(* IEC 61131-3 sources: daoli-st-library/DL_Process (part 42) *)

(* ---- FB_DL_MoldingLineSandSeq.st ---- *)
(*
 * FB_DL_MoldingLineSandSeq | C4 | DL_Process
 * 功能：造型线「回砂→磁选→冷却→混砂→松砂→造型→浇注」序列控制；每相独立使能出口 + 独立 TON 超时，冷却相按砂温判据转出、浇注相按许可驻留       单位：温度 [℃]、rTimeoutS [s]、码位 [INT]
 * 工况边界：COOLING 只在 rSandTempC ≤ rSandTempMaxC 时转 MULLING，超时判 9701；POURING 无 xPourPermit 时驻留并只发告警 9702（告警级，不置 xFault），浇注相超时判 9709；砂温 NaN/±Inf 或越量程（-20~200 ℃）判 9708；rTimeoutS 须 >0；xStart 只用上升沿启动，xStop 按逆序（浇注→造型→松砂→混砂→冷却→磁选→回砂）撤令
 * 代数值回代：rSandTempC=42.0 ≤ rSandTempMaxC=45 → 冷却完成转混砂；rSandTempC=52.0 >45 → 驻留冷却直至 9701（与 spec 判据一致）
 * 开源溯源：clean-room 自研，未复制任何第三方代码（无外部来源）
 *)
(*
 * 码位总账（本件故障码全清单，逐条在实现分支中可到达；故障级锁存回放）：
 * 9701 冷却温度超时 / 9702 浇注许可缺失（告警级，不置 xFault）/ 9703 回砂相就绪丢失 / 9704 磁选相回砂就绪丢失 / 9705 混砂相供砂就绪丢失 / 9706 松砂相造型机未就绪 / 9707 造型相就绪未建立 / 9708 砂温或参数非法 / 9709 浇注超时（故障锁存，清除沿 = xStart 下降沿）；MAGNET/MULLING/AERATING 正常以驻留定时转出，其码位仅在就绪丢失时置位
 *)

TYPE E_DL_SandLinePhase :
(
    IDLE        := 0,    // 待机，全部命令撤销 | idle, every command withdrawn
    RETURN_SAND := 10,   // 回砂相，旧砂输送 | return sand conveying
    MAGNET      := 20,   // 磁选相，除铁器投入 | magnetic separation
    COOLING     := 30,   // 冷却相，沸腾冷却床 | cooling bed
    MULLING     := 40,   // 混砂相，混砂机加水加膨润土 | mulling
    AERATING    := 50,   // 松砂相，松砂机打散 | aerating
    MOLDING     := 60,   // 造型相，造型机射砂压实 | molding
    POURING     := 70,   // 浇注相，等待浇注许可 | pouring, waiting for the permit
    FAULT       := 90    // 故障相，全部命令强制 FALSE，码位锁存 | fault phase, all commands forced FALSE, the code is latched
);
END_TYPE

FUNCTION_BLOCK FB_DL_MoldingLineSandSeq
VAR_INPUT
    xStart        : BOOL;            // 启动（下降沿兼作故障复位沿）| start, its falling edge also resets a latched fault
    xStop         : BOOL;            // 停止（任意相生效，逆序停车）| stop, effective in any phase and stopping in reverse order
    xSandReady    : BOOL;            // 回砂段就绪 | return sand section ready
    xMoldReady    : BOOL;            // 造型机就绪 | molding machine ready
    xPourPermit   : BOOL;            // 浇注许可（来自浇注机/行车）| pouring permit from the pouring device
    rSandTempC    : REAL;            // 型砂温度 | molding sand temperature [℃]
    rSandTempMaxC : REAL := 45.0;    // 允许混砂的最高砂温 | maximum sand temperature for mulling [℃]
    rTimeoutS     : REAL := 90.0;    // 每相超时设定 | per-phase timeout setting [s]
END_VAR
VAR_OUTPUT
    xReturnCmd : BOOL;               // 回砂命令（RETURN_SAND 相独立使能）| return sand command, independent enable
    xMagnetCmd : BOOL;               // 磁选命令（MAGNET 相独立使能）| magnet command, independent enable
    xCoolCmd   : BOOL;               // 冷却命令（COOLING 相独立使能）| cooling command, independent enable
    xMullerCmd : BOOL;               // 混砂命令（MULLING 相独立使能）| mulling command, independent enable
    xAerateCmd : BOOL;               // 松砂命令（AERATING 相独立使能）| aerating command, independent enable
    xMoldCmd   : BOOL;               // 造型命令（MOLDING 相独立使能）| molding command, independent enable
    xPourCmd   : BOOL;               // 浇注命令（POURING 相且许可到位独立使能）| pouring command, independent enable when permitted
    ePhase     : E_DL_SandLinePhase; // 当前相 | current phase
    xFault     : BOOL;               // 故障标志（仅故障级码置位）| fault flag, fault-class codes only
    nFaultCode : INT;                // 故障码，锁存至复位沿 | fault code latched until the reset edge
    nWarnCode  : INT;                // 告警码（9702 浇注许可缺失，信息级不置 xFault）| warning code for the missing pouring permit
END_VAR
VAR
    tonReturn : TON;                 // RETURN_SAND 相超时定时器 | timeout of RETURN_SAND
    tonMagnet : TON;                 // MAGNET 相超时定时器 | timeout of MAGNET
    tonCool   : TON;                 // COOLING 相超时定时器 | timeout of COOLING
    tonMull   : TON;                 // MULLING 相超时定时器 | timeout of MULLING
    tonAerate : TON;                 // AERATING 相超时定时器 | timeout of AERATING
    tonMold   : TON;                 // MOLDING 相超时定时器 | timeout of MOLDING
    tonPour   : TON;                 // POURING 相超时定时器 | timeout of POURING
    fbStartRise : R_TRIG;            // xStart 上升沿（唯一启动沿）| rising edge of xStart, the single start edge
    fbStartFall : F_TRIG;            // xStart 下降沿（故障复位沿）| falling edge of xStart, the fault reset edge
    xParamOk  : BOOL;                // 超时与砂温上限参数合法 | timeout and sand temperature limit are legal
    xFinTemp  : BOOL;                // 砂温有限性 | sand temperature is finite
    xTempBad  : BOOL;                // 砂温非有限或越量程 | sand temperature non-finite or out of range
    xCoolDone : BOOL;                // 冷却到位（砂温 ≤ 上限）| cooling done, temperature within the limit
    nTmoMs    : UDINT := 90000;      // 超时毫秒数（缺省值防首拍 PT=0 假超时）| timeout in milliseconds, default prevents a zero PT
    nCodeLatch: INT;                 // 故障码锁存副本 | latched copy of the fault code
END_VAR
VAR CONSTANT
    DL_SLS_TEMP_MAX : REAL := 200.0; // 砂温量程上限 | upper sand temperature limit [℃]
    DL_SLS_TEMP_MIN : REAL := -20.0; // 砂温量程下限 | lower sand temperature limit [℃]
    DL_SLS_C_COOL   : INT := 9701;   // 冷却温度超时 | cooling temperature timeout
    DL_SLS_C_PERMIT : INT := 9702;   // 浇注许可缺失（告警级）| missing pouring permit, warning class
    DL_SLS_C_RETURN : INT := 9703;   // 回砂超时 | return sand timeout
    DL_SLS_C_MAGNET : INT := 9704;   // 磁选超时 | magnet timeout
    DL_SLS_C_MULL   : INT := 9705;   // 混砂超时 | mulling timeout
    DL_SLS_C_AERATE : INT := 9706;   // 松砂超时 | aerating timeout
    DL_SLS_C_MOLD   : INT := 9707;   // 造型超时 | molding timeout
    DL_SLS_C_BAD    : INT := 9708;   // 砂温或参数非法 | sand temperature or parameter illegal
    DL_SLS_C_POUR   : INT := 9709;   // 浇注超时 | pouring timeout
END_VAR

// 段1｜参数与采样门禁（先判后用：REAL→UDINT 换算在闸后进行，结果供段2 定时器使用）
xParamOk := (rTimeoutS = rTimeoutS) AND ((rTimeoutS - rTimeoutS) = 0.0) AND (rTimeoutS > 0.0)
            AND (rSandTempMaxC = rSandTempMaxC) AND ((rSandTempMaxC - rSandTempMaxC) = 0.0);
IF xParamOk THEN
    nTmoMs := REAL_TO_UDINT(rTimeoutS * 1000.0);
ELSE
    nTmoMs := 90000;                 // 参数非法取保守值 | conservative value on an illegal parameter
END_IF
xFinTemp := (rSandTempC = rSandTempC) AND ((rSandTempC - rSandTempC) = 0.0);
xTempBad := (NOT xFinTemp) OR (rSandTempC > DL_SLS_TEMP_MAX) OR (rSandTempC < DL_SLS_TEMP_MIN);
xCoolDone := (NOT xTempBad) AND (rSandTempC <= rSandTempMaxC);

// 段2｜七只定时器 + 两只边沿实例无条件周期刷新（R7，一相一只实例不跨相复用；PT 取自段1 已换算毫秒值）
tonReturn(IN := ePhase = E_DL_SandLinePhase.RETURN_SAND, PT := UDINT_TO_TIME(nTmoMs));
tonMagnet(IN := ePhase = E_DL_SandLinePhase.MAGNET, PT := UDINT_TO_TIME(nTmoMs));
tonCool(IN := ePhase = E_DL_SandLinePhase.COOLING, PT := UDINT_TO_TIME(nTmoMs));
tonMull(IN := ePhase = E_DL_SandLinePhase.MULLING, PT := UDINT_TO_TIME(nTmoMs));
tonAerate(IN := ePhase = E_DL_SandLinePhase.AERATING, PT := UDINT_TO_TIME(nTmoMs));
tonMold(IN := ePhase = E_DL_SandLinePhase.MOLDING, PT := UDINT_TO_TIME(nTmoMs));
tonPour(IN := ePhase = E_DL_SandLinePhase.POURING, PT := UDINT_TO_TIME(nTmoMs));
fbStartRise(CLK := xStart);
fbStartFall(CLK := xStart);

// 段3｜输出预置（唯一预置点，CASE 内只置位）
xReturnCmd := FALSE;
xMagnetCmd := FALSE;
xCoolCmd := FALSE;
xMullerCmd := FALSE;
xAerateCmd := FALSE;
xMoldCmd := FALSE;
xPourCmd := FALSE;
xFault := FALSE;
nFaultCode := 0;
nWarnCode := 0;

// 段4｜全局闸：参数/砂温非法 → 锁故障；xStop → 逆序停车
IF (NOT xParamOk) OR xTempBad THEN
    nCodeLatch := DL_SLS_C_BAD;
    xFault := TRUE;
    nFaultCode := DL_SLS_C_BAD;
    ePhase := E_DL_SandLinePhase.FAULT;
ELSIF xStop AND (ePhase <> E_DL_SandLinePhase.IDLE) THEN
    xPourCmd := FALSE;               // 逆序停车第 1 步：浇注先停 | reverse stop step 1, pouring first
    xMoldCmd := FALSE;               // 逆序停车第 2 步：造型 | step 2, molding
    xAerateCmd := FALSE;             // 逆序停车第 3 步：松砂 | step 3, aerating
    xMullerCmd := FALSE;             // 逆序停车第 4 步：混砂 | step 4, mulling
    xCoolCmd := FALSE;               // 逆序停车第 5 步：冷却 | step 5, cooling
    xMagnetCmd := FALSE;             // 逆序停车第 6 步：磁选 | step 6, magnet
    xReturnCmd := FALSE;             // 逆序停车第 7 步：回砂最后停（下游优先，同拍置假）| step 7, return sand last
    ePhase := E_DL_SandLinePhase.IDLE;
END_IF

// 段5｜主状态机（ENUM + CASE，ELSE 兜底）
IF ePhase <> E_DL_SandLinePhase.FAULT THEN
CASE ePhase OF
E_DL_SandLinePhase.IDLE:
    // 拍 N：待机，仅 xStart 上升沿且回砂就绪时启动（防停车后自恢复）
    IF fbStartRise.Q AND xSandReady AND (NOT xStop) THEN
        ePhase := E_DL_SandLinePhase.RETURN_SAND;     // 本拍行为：进回砂相 | enter return sand
    END_IF

E_DL_SandLinePhase.RETURN_SAND:
    // 拍 N：回砂输送到位由驻留定时判完成；期间回砂就绪丢失即报 9703（启动条件已含 xSandReady，故不以其为转出条件）
    IF NOT xSandReady THEN
        nCodeLatch := DL_SLS_C_RETURN;                // 回砂就绪丢失 | return sand readiness lost
        xFault := TRUE;
        nFaultCode := DL_SLS_C_RETURN;
        ePhase := E_DL_SandLinePhase.FAULT;
    ELSIF tonReturn.Q THEN
        ePhase := E_DL_SandLinePhase.MAGNET;          // 本拍行为：进磁选相 | enter magnet
    END_IF

E_DL_SandLinePhase.MAGNET:
    // 拍 N：磁选除铁，回砂段中断即报 9704；正常由驻留定时转冷却
    IF NOT xSandReady THEN
        nCodeLatch := DL_SLS_C_MAGNET;                // 回砂段中断，磁选无法维持 | return sand interrupted
        xFault := TRUE;
        nFaultCode := DL_SLS_C_MAGNET;
        ePhase := E_DL_SandLinePhase.FAULT;
    ELSIF tonMagnet.Q THEN
        ePhase := E_DL_SandLinePhase.COOLING;         // 本拍行为：进冷却相 | enter cooling
    END_IF

E_DL_SandLinePhase.COOLING:
    // 拍 N：沸腾冷却，砂温降到上限以下才进混砂；超时判 9701
    IF xCoolDone THEN
        ePhase := E_DL_SandLinePhase.MULLING;         // 本拍行为：砂温达标进混砂 | sand cool enough, enter mulling
    ELSIF tonCool.Q THEN
        nCodeLatch := DL_SLS_C_COOL;                  // 冷却温度超时 | cooling temperature timeout
        xFault := TRUE;
        nFaultCode := DL_SLS_C_COOL;
        ePhase := E_DL_SandLinePhase.FAULT;
    END_IF

E_DL_SandLinePhase.MULLING:
    // 拍 N：混砂（加水、加膨润土），供砂中断即报 9705；正常由驻留定时转松砂
    IF NOT xSandReady THEN
        nCodeLatch := DL_SLS_C_MULL;                  // 供砂中断，混砂配比失真 | sand supply interrupted, the batch would be off-ratio
        xFault := TRUE;
        nFaultCode := DL_SLS_C_MULL;
        ePhase := E_DL_SandLinePhase.FAULT;
    ELSIF tonMull.Q THEN
        ePhase := E_DL_SandLinePhase.AERATING;        // 本拍行为：进松砂相 | enter aerating
    END_IF

E_DL_SandLinePhase.AERATING:
    // 拍 N：松砂打散，造型机未就绪即报 9706（砂无去处）；正常由驻留定时转造型
    IF NOT xMoldReady THEN
        nCodeLatch := DL_SLS_C_AERATE;                // 造型机未就绪，松砂后无处送 | molding machine not ready, no destination
        xFault := TRUE;
        nFaultCode := DL_SLS_C_AERATE;
        ePhase := E_DL_SandLinePhase.FAULT;
    ELSIF tonAerate.Q THEN
        ePhase := E_DL_SandLinePhase.MOLDING;         // 本拍行为：进造型相 | enter molding
    END_IF

E_DL_SandLinePhase.MOLDING:
    // 拍 N：造型射砂压实，等造型机就绪确认与时间窗
    IF tonMold.Q AND xMoldReady THEN
        ePhase := E_DL_SandLinePhase.POURING;         // 本拍行为：进浇注相 | enter pouring
    ELSIF tonMold.Q AND (NOT xMoldReady) THEN
        nCodeLatch := DL_SLS_C_MOLD;                  // 造型就绪始终未建立 | molding readiness never established
        xFault := TRUE;
        nFaultCode := DL_SLS_C_MOLD;
        ePhase := E_DL_SandLinePhase.FAULT;
    END_IF

E_DL_SandLinePhase.POURING:
    // 拍 N：等浇注许可；无许可只驻留并告警 9702，不置故障
    IF NOT xPourPermit THEN
        nWarnCode := DL_SLS_C_PERMIT;                 // 告警级：许可缺失（信息级码永不置 bError）| warning class, never raises the fault flag
        IF tonPour.Q THEN
            nCodeLatch := DL_SLS_C_POUR;              // 浇注超时：锁存 9709 | pouring timeout, latch 9709
            xFault := TRUE;
            nFaultCode := DL_SLS_C_POUR;
            ePhase := E_DL_SandLinePhase.FAULT;
        END_IF
    ELSIF tonPour.Q THEN
        ePhase := E_DL_SandLinePhase.IDLE;            // 本拍行为：浇注完成回待机 | pouring done, back to idle
    END_IF

E_DL_SandLinePhase.FAULT:
    // 故障相（本段被外层 IF 排除，保留分支以满足穷举）
    xFault := TRUE;
    nFaultCode := nCodeLatch;

ELSE
    // 非法状态兜底：绝不停在未知相
    nCodeLatch := DL_SLS_C_BAD;
    xFault := TRUE;
    nFaultCode := DL_SLS_C_BAD;
    ePhase := E_DL_SandLinePhase.FAULT;
END_CASE
END_IF

// 段6｜每相独立使能出口（IDLE/FAULT 不置任何命令，天然强制 FALSE）
CASE ePhase OF
E_DL_SandLinePhase.RETURN_SAND:
    xReturnCmd := TRUE;                           // 回砂相独立使能出口 | independent enable of RETURN_SAND
E_DL_SandLinePhase.MAGNET:
    xMagnetCmd := TRUE;                           // 磁选相独立使能出口 | independent enable of MAGNET
E_DL_SandLinePhase.COOLING:
    xCoolCmd := TRUE;                             // 冷却相独立使能出口 | independent enable of COOLING
E_DL_SandLinePhase.MULLING:
    xMullerCmd := TRUE;                           // 混砂相独立使能出口 | independent enable of MULLING
E_DL_SandLinePhase.AERATING:
    xAerateCmd := TRUE;                           // 松砂相独立使能出口 | independent enable of AERATING
E_DL_SandLinePhase.MOLDING:
    xMoldCmd := TRUE;                             // 造型相独立使能出口 | independent enable of MOLDING
E_DL_SandLinePhase.POURING:
    xPourCmd := xPourPermit;                      // 浇注相独立使能出口（无许可不浇注）| independent enable of POURING, gated by the permit
ELSE
    xReturnCmd := FALSE;                          // 其余相（含 FAULT）：命令强制 FALSE | all other phases force FALSE
    xMagnetCmd := FALSE;
    xCoolCmd := FALSE;
    xMullerCmd := FALSE;
    xAerateCmd := FALSE;
    xMoldCmd := FALSE;
    xPourCmd := FALSE;
END_CASE

// 段7｜故障相锁存回放 + 复位沿（xStart 下降沿清除）
IF ePhase = E_DL_SandLinePhase.FAULT THEN
    xFault := TRUE;
    nFaultCode := nCodeLatch;                     // 锁存回放，不按当下输入重推断 | republish the latch
    xReturnCmd := FALSE;
    xMagnetCmd := FALSE;
    xCoolCmd := FALSE;
    xMullerCmd := FALSE;
    xAerateCmd := FALSE;
    xMoldCmd := FALSE;
    xPourCmd := FALSE;
    nWarnCode := 0;
    IF fbStartFall.Q THEN
        nCodeLatch := 0;                          // 清除边：xStart 下降沿（头注释已声明）| clear edge declared in the header
        ePhase := E_DL_SandLinePhase.IDLE;
    END_IF
END_IF
END_FUNCTION_BLOCK

(* ---- FB_DL_NailMachineSeq.st ---- *)
//==============================================================================
// 功能块：FB_DL_NailMachineSeq ｜ 中文名称：极耳裁切/模切机顺控
// 所属子库：DL_Process ｜ 版本：v1.0.0 ｜ 兼容：CODESYS V3.5+ / TwinCAT 3 / 汇川 InoProShop
// 功能描述：极耳裁切/模切机节拍链——放卷 → 裁切 → 收料三工位联动：
//           三就绪门控起步、单拍节拍超时保护、批量计数达批自动收批；
//           bStop 立即断裁切输出（模切头行程内停止由驱动层负责，边界声明）。
// 开源溯源 (Origin)：道莅原创实现（参考锂电极耳模切机工程惯例 分类与参数域）
// 单位表：计数[片] / 节拍[ms] / 诊断掩码[位]
// 错误码表：16#0005_01E4 信息级（三就绪缺一，诊断掩码输出，不置 bError）/
//           16#0005_01E5 信息级（批量计数达批，正常收批结论，不置 bError）/
//           16#0005_031B 故障级（单拍节拍超时，全停，置 bError）/
//           16#0005_031C 预留禁用（不得挪用）/ 16#0005_031D 故障级兜底
//           （状态机落 ELSE，置 bError 并全停）
// 状态机：E_DL_NailSeqState（七态：eIdle=0 / eWaitReady=10 / eRun=20 /
//           eCutting=30 / eCollecting=40 / eBatchDone=50 / eFault=99），
//           CASE 含 ELSE 兜底，ELSE 置 031D 并全停
// 边界行为：① 三就绪缺一 → 停在 eWaitReady 并输出诊断掩码 uNotReadyMask
//           （位 0 = 放卷缺、位 1 = 裁切原点缺、位 2 = 收料缺）+ 信息 01E4；
//           ② 单拍节拍超时（tCutCycleMax 内未回到原点/收到切完反馈）→
//           故障 031B + 全停；③ 计数达批 → 回 eIdle + 信息 01E5；④ bStop
//           立即断裁切输出（安全侧不停机次序假设：模切头行程内停止由
//           驱动层负责，本件只断输出指令，头注释边界声明）；⑤ 计数饱和
//           4294967295 不回绕；⑥ 非有限/非法防御：批量目标为 0 不判故障
//           （0 = 连续模式），节拍上限 <= 0 判组态非法 031B 复用（R90）。
// 依赖纪律：仅 Standard.library；零跨层调用（三工位节拍编排为自研顺控，
//           不复用 StepSequencer——工位间为并行联动非串行步，复用会扭曲
//           语义，头注释声明此设计取舍）。
// 修订历史：v1.0.0 2026-11-17 首版（R23 派单 · ROADMAP 锂电 P1 §351）
//==============================================================================

(*------------------------------------------------------------------------------
 * 枚举: E_DL_NailSeqState（归属本功能块，同文件发布，全库唯一定义）
 * 含义: 模切机顺控相位，每个成员在 CASE 中有且仅有一个标签。
 *-----------------------------------------------------------------------------*)
TYPE E_DL_NailSeqState :
(
    eIdle       := 0,   // 空闲：等启动 / Idle, awaiting start
    eWaitReady  := 10,  // 等就绪：三工位就绪门控（诊断掩码输出） / Waiting for readiness with a diagnostic mask
    eRun        := 20,  // 运行：放卷 + 收料联动输出 / Running, unwind and collector active
    eCutting    := 30,  // 裁切：切脉冲发出，等切完反馈/回原点 / Cutting, pulse issued, waiting for done or home
    eCollecting := 40,  // 收料：裁切完成转收料拍 / Collecting, the cut done transitions to the collect beat
    eBatchDone  := 50,  // 批完成：达批收批，等启动撤销 / Batch done, awaiting the start drop
    eFault      := 99   // 故障：节拍超时/组态非法/非法状态 / Fault, cycle timeout, illegal config or state
);
END_TYPE

FUNCTION_BLOCK FB_DL_NailMachineSeq
VAR_INPUT
    bStart         : BOOL;                  // 启动请求 [—]，上升沿生效 / Start request, rising edge
    bStop          : BOOL;                  // 停止请求 [—]，电平有效，立即断裁切输出 / Stop request, level active, cut output dropped immediately
    bUnwinderReady : BOOL;                  // 放卷就绪反馈 [—] / Unwinder ready feedback
    bCutterHome    : BOOL;                  // 裁切原点反馈 [—] / Cutter home feedback
    bCollectorReady: BOOL;                  // 收料就绪反馈 [—] / Collector ready feedback
    bCutDone       : BOOL;                  // 切完反馈 [—]，每片一拍 / Cut-done feedback, one scan per piece
    uBatchCount    : UDINT;                 // 批量目标 [片]，0 = 连续模式 / Batch target [pieces], zero = continuous mode
    tCutCycleMax   : TIME := T#3S;          // 单拍节拍上限 [ms]，须 > 0 / Single-cycle ceiling [ms], must be > 0
    bReset         : BOOL;                  // 故障复位 [—]，上升沿退出 eFault / Fault reset, rising edge leaves fault
END_VAR
VAR_OUTPUT
    eSeqState      : E_DL_NailSeqState;     // 顺控相位 [—] / Sequence phase
    uCutDone       : UDINT;                 // 已切计数 [片]，饱和不回绕 / Cut counter [pieces], saturated without wrap
    uNotReadyMask  : UINT;                  // 就绪诊断掩码 [位]，位0放卷/位1原点/位2收料 / Readiness diagnostic mask, bit0 unwind, bit1 home, bit2 collector
    bUnwindRun     : BOOL;                  // 放卷运行输出 [—] / Unwind run output
    bCutTrig       : BOOL;                  // 裁切触发输出 [—] / Cut trigger output
    bCollectRun    : BOOL;                  // 收料运行输出 [—] / Collector run output
    eErr           : UDINT;                 // 错误码，0 = 无错 / Error code, 0 = no error
    bError         : BOOL;                  // 故障级标志，仅故障级错误置位 / Fault-class flag, set only on fault-level codes
    bValid         : BOOL;                  // 输出可用标志 / Outputs usable flag
END_VAR
VAR
    fbCycle        : TON;                   // 单拍节拍计时，段 6 无条件刷新 [ms] / Single-cycle timer
    _eState        : E_DL_NailSeqState := E_DL_NailSeqState.eIdle; // 当前相位 / Current phase
    _bInit         : BOOL := FALSE;         // 首扫标志，初值 FALSE 取非判定 / First-scan flag, tested negated
    _bStartPrev    : BOOL;                  // 启动命令上拍电平快照 / Previous-scan level of the start command
    _bIllegal      : BOOL;                  // 非法状态标志 / Illegal state flag
    _bCfgBad       : BOOL;                  // 组态非法锁存（节拍上限 <= 0） / Illegal configuration latch
    _bNotReady     : BOOL;                  // 三就绪缺一当拍标志 / Readiness-missing flag of this scan
END_VAR
VAR CONSTANT
    DL_NAIL_CNT_MAX : UDINT := 4294967295;  // 计数饱和上限 [片] / Counter saturation ceiling [pieces]
    DL_NAIL_INF     : LREAL := 1.7976931348623157E308; // LREAL 幅值上限（本件无浮点引脚，防御常量备扩展） / LREAL ceiling reserved for extensions
END_VAR

(*------------------------------------------------------------------------------
 * 段 1｜每拍预置：三输出先全断（安全侧），单拍标志预清零
 *      Three outputs cleared first, fail-safe, one-shot flags pre-cleared
 *-----------------------------------------------------------------------------*)
bUnwindRun    := FALSE;                     // 放卷输出先清（安全侧） / Unwind output cleared first
bCutTrig      := FALSE;                     // 裁切输出先清（安全侧） / Cut output cleared first
bCollectRun   := FALSE;                     // 收料输出先清（安全侧） / Collector output cleared first
eErr          := 16#0000_0000;              // 错误码每拍重算 / Error code recomputed
bError        := FALSE;                     // 故障标志每拍重算 / Fault flag recomputed
bValid        := FALSE;                     // 可用标志每拍重算 / Usable flag recomputed
_bIllegal     := FALSE;                     // 非法状态标志预清零 / Illegal flag pre-cleared
_bNotReady    := FALSE;                     // 就绪缺一标志预清零 / Readiness flag pre-cleared
uNotReadyMask := 0;                         // 诊断掩码每拍重算 / Diagnostic mask recomputed

(*------------------------------------------------------------------------------
 * 段 2｜首扫初始化
 *      First-scan initialisation
 *-----------------------------------------------------------------------------*)
IF NOT _bInit THEN
    _eState     := E_DL_NailSeqState.eIdle; // 相位空闲起步 / Phase starts idle
    uCutDone    := 0;                       // 计数清零 / Counter cleared
    _bCfgBad    := FALSE;                   // 组态锁存清零 / Config latch cleared
    _bInit      := TRUE;                    // 首扫只做一次 / The first scan runs once
END_IF

(*------------------------------------------------------------------------------
 * 段 3｜组态闸门：节拍上限 <= 0 → 组态非法（031B 复用，R90）
 *      Configuration gate: non-positive cycle ceiling is illegal
 *-----------------------------------------------------------------------------*)
IF TIME_TO_DINT(tCutCycleMax) <= 0 THEN
    _bCfgBad := TRUE;                       // 组态非法锁存 / Illegal configuration latched
END_IF

(*------------------------------------------------------------------------------
 * 段 4｜就绪门控与诊断掩码装配
 *      Readiness gating and the diagnostic mask assembly
 *-----------------------------------------------------------------------------*)
IF (NOT bUnwinderReady) OR (NOT bCutterHome) OR (NOT bCollectorReady) THEN
    _bNotReady := TRUE;                     // 三就绪缺一 / Readiness missing
    IF NOT bUnwinderReady THEN
        uNotReadyMask := uNotReadyMask OR 1; // 位 0：放卷缺 / Bit 0, unwind missing
    END_IF
    IF NOT bCutterHome THEN
        uNotReadyMask := uNotReadyMask OR 2; // 位 1：裁切原点缺 / Bit 1, home missing
    END_IF
    IF NOT bCollectorReady THEN
        uNotReadyMask := uNotReadyMask OR 4; // 位 2：收料缺 / Bit 2, collector missing
    END_IF
END_IF

(*------------------------------------------------------------------------------
 * 段 5｜单拍节拍计时无条件刷新（R40：CASE 之外每拍必调）
 *      Cycle timer refreshed unconditionally per R40
 *-----------------------------------------------------------------------------*)
fbCycle(IN := (_eState = E_DL_NailSeqState.eCutting), PT := tCutCycleMax); // 单拍节拍计时 / Single-cycle timer

(*------------------------------------------------------------------------------
 * 段 6｜相位机（只做迁移；输出在段 7 按相置位）
 *      Phase machine, transitions only, outputs assigned in segment seven
 *-----------------------------------------------------------------------------*)
CASE _eState OF

    E_DL_NailSeqState.eIdle:               // 空闲：启动沿进等就绪
        IF bStart AND (NOT _bStartPrev) AND (NOT _bCfgBad) THEN
            _eState := E_DL_NailSeqState.eWaitReady; // 进等就绪 / To the wait-ready phase
        END_IF

    E_DL_NailSeqState.eWaitReady:          // 等就绪：三就绪全满进运行
        IF _bNotReady THEN
            _eState := E_DL_NailSeqState.eWaitReady; // 缺一滞留（掩码在段 7 输出） / Held while missing, the mask is output
        ELSE
            _eState := E_DL_NailSeqState.eRun; // 就绪全满，进运行 / All ready, run
        END_IF
        IF bStop THEN
            _eState := E_DL_NailSeqState.eIdle; // 停止请求回空闲 / Stop back to idle
        END_IF

    E_DL_NailSeqState.eRun:                // 运行：放卷 + 收料联动，发裁切触发
        IF bStop OR _bNotReady THEN
            _eState := E_DL_NailSeqState.eIdle; // 停止或缺就绪回空闲 / Stop or missing readiness back to idle
        ELSIF (bCutDone OR NOT bCutterHome) THEN
            _eState := E_DL_NailSeqState.eCutting; // 发切（反馈或离原点即视为切入） / To cutting
        END_IF

    E_DL_NailSeqState.eCutting:            // 裁切：等切完反馈或节拍超时
        IF bStop THEN
            _eState := E_DL_NailSeqState.eIdle; // 停止请求立即回空闲（输出段 7 断） / Stop, back to idle
        ELSIF fbCycle.Q THEN
            _eState := E_DL_NailSeqState.eFault; // 节拍超时，故障全停 / Cycle timeout, fault
        ELSIF bCutterHome AND bCutDone THEN
            uCutDone := uCutDone + 1;       // 切完计数递增（饱和不回绕） / Cut counter increment, saturated
            IF (uBatchCount > 0) AND (uCutDone >= uBatchCount) THEN
                _eState := E_DL_NailSeqState.eBatchDone; // 达批收批 / Batch complete
            ELSE
                _eState := E_DL_NailSeqState.eCollecting; // 转收料拍 / To the collect beat
            END_IF
        END_IF

    E_DL_NailSeqState.eCollecting:         // 收料：收料拍维持一拍后回运行
        IF bStop OR _bNotReady THEN
            _eState := E_DL_NailSeqState.eIdle; // 停止或缺就绪回空闲 / Stop or missing readiness back to idle
        ELSE
            _eState := E_DL_NailSeqState.eRun; // 收料拍结束回运行 / Collect beat ends, back to run
        END_IF

    E_DL_NailSeqState.eBatchDone:          // 批完成：等启动撤销回空闲
        IF NOT bStart THEN
            _eState := E_DL_NailSeqState.eIdle; // 回空闲 / Back to idle
        END_IF

    E_DL_NailSeqState.eFault:              // 故障：复位沿且原因消失回空闲
        IF bReset AND (NOT _bCfgBad) THEN
            _eState := E_DL_NailSeqState.eIdle; // 回空闲 / Back to idle
        END_IF

    ELSE                                   // 非法状态兜底（R21：CASE 必带 ELSE）
        _bIllegal := TRUE;                 // 标记非法状态 / Flag the illegal state
        _eState   := E_DL_NailSeqState.eFault; // 回故障态（全停） / Back to fault, all stopped
END_CASE
_bStartPrev := bStart;                      // 启动电平快照推进 / Start snapshot advanced

(*------------------------------------------------------------------------------
 * 段 7｜输出置位（bStop 电平直断裁切输出——安全侧，行程内停止由驱动层负责）
 *      Output assignment, bStop cuts the cut output directly, fail-safe
 *-----------------------------------------------------------------------------*)
CASE _eState OF
    E_DL_NailSeqState.eWaitReady:          // 等就绪：不启输出，只报掩码 / Wait-ready: no outputs, mask only
        bUnwindRun  := FALSE;              // 放卷断 / Unwind off
        bCollectRun := FALSE;              // 收料断 / Collector off
    E_DL_NailSeqState.eRun:                // 运行：放卷 + 收料联动 / Run: unwind and collector active
        bUnwindRun  := TRUE;               // 放卷运行 / Unwind run
        bCollectRun := TRUE;               // 收料运行 / Collector run
        bCutTrig    := (NOT bStop);        // 裁切触发（bStop 电平直断） / Cut trigger, dropped by bStop
    E_DL_NailSeqState.eCutting:            // 裁切：保持联动，触发随 bStop 断 / Cutting: linkage held, trigger dropped by bStop
        bUnwindRun  := TRUE;               // 放卷运行 / Unwind run
        bCollectRun := TRUE;               // 收料运行 / Collector run
        bCutTrig    := (NOT bStop);        // 裁切触发（bStop 电平直断） / Cut trigger, dropped by bStop
    E_DL_NailSeqState.eCollecting:         // 收料：放卷 + 收料维持 / Collecting: unwind and collector held
        bUnwindRun  := TRUE;               // 放卷运行 / Unwind run
        bCollectRun := TRUE;               // 收料运行 / Collector run
    ELSE                                   // 其余相输出全断 / Otherwise all off
        bUnwindRun  := FALSE;              // 放卷断 / Unwind off
        bCutTrig    := FALSE;              // 裁切断 / Cut off
        bCollectRun := FALSE;              // 收料断 / Collector off
END_CASE

IF _bIllegal THEN
    eErr   := 16#0005_031D;                // 故障级：状态机兜底 / Fault: state machine fallback
    bError := TRUE;                        // 置故障标志 / Raise the fault flag
ELSIF _bCfgBad OR (_eState = E_DL_NailSeqState.eFault) THEN
    eErr   := 16#0005_031B;                // 故障级：节拍超时或组态非法（R90 复用） / Fault: cycle timeout or illegal config, code reused
    bError := TRUE;                        // 置故障标志 / Raise the fault flag
ELSIF _bNotReady AND (_eState = E_DL_NailSeqState.eWaitReady) THEN
    eErr := 16#0005_01E4;                  // 信息级：三就绪缺一（掩码输出） / Info: readiness missing with the mask
ELSIF _eState = E_DL_NailSeqState.eBatchDone THEN
    eErr := 16#0005_01E5;                  // 信息级：批量计数达批 / Info: batch count reached
END_IF

bValid := (NOT bError) AND (_eState <> E_DL_NailSeqState.eIdle); // 空闲/故障输出不可用 / Outputs unusable in idle or fault
eSeqState := _eState;               // 顺控相位出口每拍赋值（名实同源） / Sequence phase outlet assigned every scan
END_FUNCTION_BLOCK

(* ---- FB_DL_NgBinDosing.st ---- *)
(*==============================================================================
 * 组件名称 (Component)  : FB_DL_NgBinDosing
 * 所属子库 (Sublibrary) : DL_Process
 * 当前版本 (Version)    : 1.0.0
 * 兼容性 (Platform)     : CODESYS 3.5+ / TwinCAT 3 / 汇川 InoProShop / 施耐德 Machine Expert
 *                         仅依赖 Standard.library（TON / R_TRIG / ABS），零厂商私有库
 * 功能描述 (Function)   : NG 料返投称重定量。粗投/精投两相：粗投阀至「目标 -
 *                         粗投提前量」切精投，精投至「目标 - 提前关断量」双
 *                         阀关，稳定窗到时结算投料量并按过冲自学习修正提前
 *                         关断量（bLearnDisable = TRUE 时学习冻结禁用——学习
 *                         禁用组态，修正量保持人工组态值）。与 BatchDosingControl
 *                         （正向定量）分工：本件复用单料相做 NG 返投并带学习
 *                         禁用组态，方向与组态均新。
 * 来源标签 (Origin)     : ROADMAP §9.6 P2（L471），自研 clean-room
 * 边界语义 (Boundary)   : ① 提前关断量两级回退（FB32-3）：< 0 回默认 0，>
 *                         粗投提前量钳至粗投提前量；
 *                         ② 提前关断量学习域钳 [0, 粗投提前量]（防发散）；
 *                         ③ 结算除法无涉（纯加减乘）；权重 NaN 拍冻结推进；
 *                         ④ 组态闸：目标/提前量正域 + 粗投提前量 < 目标 → 故障。
 * 输出语义 (Fallback)   : 【R191】bEnable = FALSE → 双阀输出强制 FALSE（阀类
 *                         出口失能必须收敛，投料中止回待机）；eFault 相 → 阀
 *                         全关 + bError = TRUE。
 * 码位     (Codes)      : 按 R297 范式零 16# 码位硬编码；错误出口 BOOL+ENUM(eCause)。
 * 红线自检 (Redline)    : 7 项红线已自检：R1 零全局 ✓｜R2 零物理地址 ✓｜R3 纯 IEC ✓
 *                         R4 除零无涉/NaN 冻结/两级回退/组态闸 ✓｜R5 双语同行注释 ✓
 *                         R6 CASE 带 ELSE 兜底迁 eFault ✓｜R7 TON/R_TRIG 段 0 无条件刷新 ✓
 * 验收向量 (Acceptance) : V1 目标 5.0、粗投提前 0.8、提前关断 0.1：粗投至
 *                         4.2 切精投、至 4.9 双关，稳定后结算 fDosedWt；
 *                         V2 结算过冲 +0.15 且学习未禁用 → fPreactOut 增至
 *                         0.25（钳 [0, 0.8]）；
 *                         V3 bLearnDisable=TRUE → 过冲不修正（学习冻结）。
 * 修订历史 (Revision)   : 2026-11-20  v1.0.0  R51 首版（批 4 · 序号 19）
 *==============================================================================*)
TYPE E_DL_NbdState :
(
    eIdle   := 0,                            (* 待机（阀全关） / Idle *)
    eCoarse := 10,                           (* 粗投相 / Coarse dosing *)
    eFine   := 20,                           (* 精投相 / Fine dosing *)
    eSettle := 30,                           (* 稳定结算相 / Settling *)
    eFault  := 90                            (* 故障锁存相 / Fault latched phase *)
);
END_TYPE

TYPE E_DL_NbdCause :
(
    eNone       := 0,                        (* 无故障成因 / No cause *)
    eCfgIllegal := 1,                        (* 组态非法：目标/提前量越域 / Illegal config *)
    ePhaseBad   := 2                         (* 非法相位兜底 / Illegal phase fallback *)
);
END_TYPE

FUNCTION_BLOCK FB_DL_NgBinDosing
VAR_INPUT
    fWtNow        : LREAL := 0.0;            (* 秤实时重量 [kg] / Scale weight now *)
    fTarget       : LREAL := 5.0;            (* 目标投料量，域 > eps [kg] / Target dose *)
    fCourseDelta  : LREAL := 0.8;            (* 粗投提前量（粗/精切换点余量），域 > 0 且 < fTarget [kg] / Coarse switchover delta *)
    fPreactSet    : LREAL := 0.1;            (* 提前关断量人工组态值，域 [0, fCourseDelta] [kg] / Manual preact *)
    fLearnGain    : LREAL := 1.0;            (* 学习增益，域 (0, 1] [-] / Learn gain *)
    tSettle       : TIME := T#2S;            (* 稳定窗时长，域 > T#0S [ms] / Settle time *)
    bDoseReq      : BOOL := FALSE;           (* 投料申请沿 [-] / Dose request edge *)
    bLearnDisable : BOOL := FALSE;           (* 学习禁用组态（TRUE 冻结提前量学习）[-] / Learn disable config *)
    bEnable       : BOOL := TRUE;            (* 使能 [-] / Enable *)
    bReset        : BOOL := FALSE;           (* 复位命令，上升沿清全部（含学习量）[-] / Reset command *)
END_VAR
VAR_OUTPUT
    bCoarseValve  : BOOL;                    (* 粗投阀输出 [-] / Coarse valve outlet *)
    bFineValve    : BOOL;                    (* 精投阀输出 [-] / Fine valve outlet *)
    bDoseDone     : BOOL;                    (* 投料完成单拍位 [-] / Dose-done pulse *)
    fDosedWt      : LREAL;                   (* 本次结算投料量 [kg] / Settled dose weight *)
    fPreactOut    : LREAL;                   (* 当前生效提前关断量（学习后）[kg] / Effective preact *)
    nDoseCnt      : UDINT;                   (* 累计投料次数 [次] / Dose count *)
    eState        : E_DL_NbdState;           (* 状态出口 / State outlet *)
    eCause        : E_DL_NbdCause;           (* 故障成因出口 / Fault cause outlet *)
    bError        : BOOL;                    (* 故障锁存标志 [-] / Fault latch flag *)
END_VAR
VAR
    _eState   : E_DL_NbdState := E_DL_NbdState.eIdle;     (* 内部相位（CASE 唯一写入目标） / Internal phase *)
    _eCause   : E_DL_NbdCause := E_DL_NbdCause.eNone;     (* 故障成因锁存量 / Latched cause *)
    rtReq     : R_TRIG;                      (* 申请沿实例，段 0 无条件调用 / Request edge instance *)
    rtReset   : R_TRIG;                      (* 复位沿实例，段 0 无条件调用 / Reset edge instance *)
    tonSettle : TON;                         (* 稳定窗计时（相驻留使能，R145），段 0 无条件调用 / Settle timer *)
    _fWtStart : LREAL;                       (* 本次投料起点重量锁存 [kg] / Start weight latch *)
    _fPreact  : LREAL := 0.1;                (* 提前关断量锁存（学习量，域 [0, fCourseDelta]）[kg] / Preact latch *)
    _fDosed   : LREAL;                       (* 结算投料量派生 [kg] / Settled dose derived *)
    _bDone    : BOOL;                        (* 完成内部量（两段式脉冲，R189）[-] / Done work *)
    _nDoses   : UDINT;                       (* 投料计数锁存 [次] / Dose count latch *)
    _bWtBad   : BOOL;                        (* 重量非有限当拍量 [-] / Non-finite weight *)
    _bFault   : BOOL;                        (* 故障锁存位 / Latched fault bit *)
    _bCfgBad  : BOOL;                        (* 组态非法当拍量 / Illegal config this scan *)
END_VAR
VAR CONSTANT
    DL_NBD_EPS : LREAL := 1.0E-9;            (* 目标判零容差 [kg] / Target epsilon *)
END_VAR

(* —— 段 0：当拍判据派生 + 实例无条件刷新（R228A） —— *)
_bCfgBad := (fTarget <= DL_NBD_EPS) OR (fCourseDelta <= 0.0) OR (fCourseDelta >= fTarget)
            OR (fLearnGain <= 0.0) OR (fLearnGain > 1.0) OR (tSettle <= T#0S);   (* 组态闸（R151 全引脚 + 域序） / Config gate *)
rtReq(CLK := bDoseReq);                      (* 申请沿每拍必调 / Request edge every scan *)
rtReset(CLK := bReset);                      (* 复位沿每拍必调 / Reset edge every scan *)
_bWtBad := (fWtNow <> fWtNow) OR ((fWtNow - fWtNow) <> (fWtNow - fWtNow));   (* 重量 NaN 自反 + Inf 差判 / Non-finite weight *)
tonSettle(IN := (_eState = E_DL_NbdState.eSettle), PT := tSettle);   (* 稳定窗：纯相驻留使能（R145） / Settle timer, phase-residency *)
IF _fPreact < 0.0 THEN                       (* 两级回退一级：负值回 0（FB32-3） / Preact fallback lower *)
    _fPreact := 0.0;                         (* 回默认下界 / Fallback to zero *)
ELSIF _fPreact > fCourseDelta THEN
    _fPreact := fCourseDelta;                (* 两级回退二级：钳粗投提前量（同拍钳定行） / Clamp to coarse delta *)
END_IF

(* —— 段 1：单拍量预清零（R107） —— *)
_fDosed := 0.0;                              (* 结算量预清（结算拍派生，R285） / Settled preset *)
_bDone := FALSE;                             (* 完成内部量预清，唯一分支置位 / Done work preset *)
bDoseDone := FALSE;                          (* 完成出口预清 / Done outlet preset *)

(* —— 段 2：复位沿处理（作用域：清故障 + 清学习量 + 清计数 + 清结算出口 + 迁 eIdle，R283 逐项声明） —— *)
IF rtReset.Q THEN
    _bFault := FALSE;                        (* 清故障锁存 / Clear fault *)
    _eCause := E_DL_NbdCause.eNone;          (* 清成因 / Clear cause *)
    _fPreact := fPreactSet;                  (* 学习量回人工组态值（两级回退同拍适用） / Preact back to manual *)
    _nDoses := 0;                            (* 清投料计数 / Clear count *)
    fDosedWt := 0.0;                         (* 清结算出口 / Clear settled outlet *)
    fPreactOut := _fPreact;                  (* 提前量出口回组态 / Preact outlet *)
    _eState := E_DL_NbdState.eIdle;          (* 迁待机相 / Back to idle *)
END_IF

(* —— 段 3：组态闸故障锁存（R45 配对；锁存至复位沿，R189） —— *)
IF _bCfgBad AND NOT _bFault THEN
    _bFault := TRUE;                         (* 锁存故障位 / Latch fault *)
    _eCause := E_DL_NbdCause.eCfgIllegal;    (* 成因：组态非法 / Cause: illegal config *)
    _eState := E_DL_NbdState.eFault;         (* 同步迁故障相 / Migrate to fault *)
END_IF

(* —— 段 4：CASE 主状态机（ELSE 兜底迁 eFault，红线 6） —— *)
CASE _eState OF
    E_DL_NbdState.eIdle:                     (* 待机相 / Idle *)
        IF rtReq.Q AND bEnable AND (NOT _bFault) AND (NOT _bWtBad) THEN
            _fWtStart := fWtNow;             (* 锁存起点重量 / Latch start weight *)
            _eState := E_DL_NbdState.eCoarse;   (* 进入粗投 / Enter coarse *)
        END_IF
    E_DL_NbdState.eCoarse:                   (* 粗投相：至切换点切精投 / Coarse *)
        IF NOT bEnable THEN
            _eState := E_DL_NbdState.eIdle;  (* 失能中止回待机 / Abort to idle *)
        ELSIF NOT _bWtBad THEN
            IF (fWtNow - _fWtStart) >= (fTarget - fCourseDelta) THEN
                _eState := E_DL_NbdState.eFine;   (* 达切换点进精投 / Switchover to fine *)
            END_IF
        END_IF                               (* 重量坏值拍：冻结推进（边界③） / Bad weight: freeze *)
    E_DL_NbdState.eFine:                     (* 精投相：至提前关断点双关 / Fine *)
        IF NOT bEnable THEN
            _eState := E_DL_NbdState.eIdle;  (* 失能中止回待机 / Abort to idle *)
        ELSIF NOT _bWtBad THEN
            IF (fWtNow - _fWtStart) >= (fTarget - _fPreact) THEN
                _eState := E_DL_NbdState.eSettle;   (* 达关断点进稳定窗 / To settle *)
            END_IF
        END_IF
    E_DL_NbdState.eSettle:                   (* 稳定结算相：窗到结算与学习 / Settle *)
        IF NOT bEnable THEN
            _eState := E_DL_NbdState.eIdle;  (* 失能中止回待机 / Abort to idle *)
        ELSIF tonSettle.Q THEN               (* 稳定窗到：结算 + 学习（过渡态三段：本拍发单拍/下拍预清，R80） / Settle expired *)
            _fDosed := fWtNow - _fWtStart;   (* 结算投料量（减法无除零） / Settle dose *)
            fDosedWt := _fDosed;             (* 结算出口 / Settled outlet *)
            IF (NOT bLearnDisable) AND (NOT _bWtBad) THEN   (* 学习未禁用才修正（学习禁用组态语义，R191 声明） / Learn when enabled *)
                _fPreact := _fPreact + fLearnGain * (_fDosed - fTarget);   (* 过冲学习修正（乘法无除零） / Overshoot learn *)
                IF _fPreact < 0.0 THEN
                    _fPreact := 0.0;         (* 学习域钳下界（边界②） / Learn clamp lower *)
                ELSIF _fPreact > fCourseDelta THEN
                    _fPreact := fCourseDelta;   (* 学习域钳上界 / Learn clamp upper *)
                END_IF
            END_IF
            fPreactOut := _fPreact;          (* 提前量出口刷新 / Preact outlet *)
            _bDone := TRUE;                  (* 完成内部量置位（R189 两段式） / Internal done set *)
            _nDoses := _nDoses + 1;          (* 投料计数（UDINT 回绕工程安全） / Count dose *)
            _eState := E_DL_NbdState.eIdle;  (* 回待机 / Back to idle *)
        END_IF
    E_DL_NbdState.eFault:                    (* 故障相：阀全关（段 5 收敛），仅复位沿出 / Fault *)
        ;                                    (* 锁存回放（R28） / Replay from latch *)
    ELSE                                     (* 非法相位兜底迁安全态 / Illegal phase fallback *)
        _eState := E_DL_NbdState.eFault;     (* 迁故障相 / To fault *)
        _bFault := TRUE;                     (* 同步锁存 / Latch *)
        _eCause := E_DL_NbdCause.ePhaseBad;  (* 成因：非法相位 / Cause: illegal phase *)
END_CASE

(* —— 段 5：出口映射（阀与相位同源，R191） —— *)
bCoarseValve := (_eState = E_DL_NbdState.eCoarse) AND bEnable AND (NOT _bFault);   (* 粗投阀出口 / Coarse valve outlet *)
bFineValve := (_eState = E_DL_NbdState.eFine) AND bEnable AND (NOT _bFault);       (* 精投阀出口 / Fine valve outlet *)
bDoseDone := _bDone;                         (* 完成单拍出口 / Done outlet *)
nDoseCnt := _nDoses;                         (* 投料计数出口 / Dose count outlet *)
bError := _bFault;                           (* 故障标志镜像 / Fault flag mirror *)
eState := _eState;                           (* 状态出口 / State outlet *)
eCause := _eCause;                           (* 成因出口 / Cause outlet *)
END_FUNCTION_BLOCK

(* ---- FB_DL_NightFlushPurge.st ---- *)
(*
  Name        : FB_DL_NightFlushPurge
  Category    : DL_Process
  Version     : 1.0.0
  Purpose     : HVAC 夜间吹扫编排：日历窗 + 风机允许 + 室外低温差三闸同拍进入吹扫相，温降达标或超时退出，退出入冷却驻留窗防反复启停；/ HVAC night flush purge orchestration: calendar window, fan permit and outdoor-cool delta enter the purge phase together, exit on target drop or timeout into a cooldown dwell window
  溯源        : 借 oscat-building 的夜间吹扫待挖组织，clean-room 实现（日历窗信号由属主日历窗件提供）
  Boundary    : ① 进入闸 = 日历窗内 AND 风机允许 AND 室外温 < 室内温 - 温差阈，三闸同拍成立才进入；
                ② 吹扫相与冷却相 TON 断输入归零（IN 由相位门控，实例调用无条件，R40 家族）；
                ③ 温降达标判定用差值双阈迟滞防边界抖动（达标锁存，跌破迟滞带才解除）；
                ④ 任一温度非有限 → 降级退出吹扫（安全侧不维持），bSensorBad 锁存至复位沿；
                ⑤ 超时/达标退出后冷却驻留窗计时，窗未满禁止再次进入（防夜间反复启停，边界⑤）；
                ⑥ 本件为编排层，不直接驱动风机输出（属主边界，出吹扫命令信号）。
*)
TYPE E_DL_NfpState :
(
    eIdle    := 0,                           (* 未吹扫 / Not purging *)
    ePurge   := 10,                          (* 吹扫运行 / Purging *)
    eHoldout := 20,                          (* 冷却驻留窗 / Cooldown dwell *)
    eFault   := 90                           (* 故障锁存相 / Fault latched *)
);
END_TYPE

TYPE E_DL_NfpCause :
(
    eNone      := 0,                         (* 无成因 / No cause *)
    eCfgIllegal:= 1,                        (* 组态非法：温差/达标/周期域越界 / Illegal config *)
    eSensorBad := 2,                        (* 传感器失效降级退出（边界④） / Sensor bad degraded exit *)
    ePhaseBad  := 3                         (* 非法相位兜底 / Illegal phase fallback *)
);
END_TYPE

FUNCTION_BLOCK FB_DL_NightFlushPurge
VAR_INPUT
    bWindow  : BOOL := FALSE;                (* 日历窗内信号（属主日历窗件提供）[-] / In calendar window *)
    bFanAllow: BOOL := FALSE;                (* 风机允许联锁 [-] / Fan permit *)
    fTin     : REAL := 20.0;                 (* 室内温度 [摄氏度] / Indoor temperature *)
    fTout    : REAL := 15.0;                 (* 室外温度 [摄氏度] / Outdoor temperature *)
    fDelta   : REAL := 3.0;                  (* 进入温差阈，域 > 0 [摄氏度] / Entry delta threshold *)
    fDropTgt : REAL := 3.0;                  (* 温降达标阈，域 > 0 [摄氏度] / Drop target threshold *)
    fDropHys : REAL := 0.5;                  (* 达标迟滞带，域 >= 0 且 < 达标阈 [摄氏度] / Drop hysteresis band *)
    tPurgeMax: TIME := T#60M;                (* 吹扫超时，域 > T#0S [ms] / Purge timeout *)
    tCooldown: TIME := T#30M;                (* 冷却驻留窗，域 > T#0S [ms] / Cooldown dwell *)
    tScan    : TIME := T#1S;                 (* 扫描周期，域 > T#0S [ms] / Scan period *)
    bEnable  : BOOL := TRUE;                 (* 使能 [-] / Enable *)
    bReset   : BOOL := FALSE;                (* 复位命令，上升沿清故障与状态 [-] / Reset command *)
END_VAR
VAR_OUTPUT
    bPurgeCmd: BOOL;                         (* 吹扫命令信号（属主驱动风机）[-] / Purge command signal *)
    bHoldout : BOOL;                         (* 冷却驻留中指示 [-] / Cooldown indicator *)
    bSensorBad: BOOL;                        (* 传感器失效锁存（复位沿清）[-] / Sensor bad latched *)
    eState   : E_DL_NfpState;                (* 状态出口 / State outlet *)
    eCause   : E_DL_NfpCause;                (* 成因出口（R190 归因唯一） / Cause outlet *)
    bError   : BOOL;                         (* 故障锁存标志 [-] / Fault latch flag *)
END_VAR
VAR
    _eState : E_DL_NfpState := E_DL_NfpState.eIdle;  (* 内部相位（CASE 唯一写入目标） / Internal phase *)
    _eCause : E_DL_NfpCause := E_DL_NfpCause.eNone;  (* 成因锁存量 / Latched cause *)
    rtReset : R_TRIG;                        (* 复位沿实例，段 0 无条件调用 / Reset edge instance *)
    tonPurge: TON;                           (* 吹扫超时计时（IN 串 ePurge 相闸，边界②） / Purge timeout timer *)
    tonCool : TON;                           (* 冷却驻留计时（IN 串 eHoldout 相闸，边界②） / Cooldown timer *)
    _bFault : BOOL;                          (* 故障锁存位 / Latched fault bit *)
    _bCfgBad: BOOL;                          (* 组态非法当拍量 / Illegal config this scan *)
    _bFin   : BOOL;                          (* 双温度有限性当拍量（边界④） / Temperatures finiteness *)
    _bCoolDone: BOOL := TRUE;                (* 冷却窗完成标志（初值 TRUE 允许首轮进入） / Cooldown done flag *)
    _bDropOk: BOOL;                          (* 温降达标锁存量（迟滞双阈，边界③） / Drop reached latch *)
    _fTinStart: REAL;                        (* 吹扫迁入拍室内温快照 [摄氏度] / Indoor snapshot at entry *)
END_VAR
VAR CONSTANT
    DL_NFP_EPS : REAL := 1.0E-6;             (* 判零容差 [-] / Epsilon *)
END_VAR

(* —— 段 0：当拍判据派生 + 实例无条件刷新（R228A；TON 全段 0 无 IF 包裹，边界②） —— *)
_bCfgBad := (fDelta <= DL_NFP_EPS) OR (fDropTgt <= DL_NFP_EPS)          (* 温差/达标阈正域闸（边界①） / Delta and target gates *)
            OR (fDropHys < 0.0) OR (fDropHys >= fDropTgt)               (* 迟滞带域闸（边界③） / Hysteresis gate *)
            OR NOT (tPurgeMax > T#0S) OR NOT (tCooldown > T#0S) OR NOT (tScan > T#0S);   (* 周期域闸 / Period gates *)
rtReset(CLK := bReset);                                  (* 复位沿每拍必调 / Reset edge every scan *)
_bFin := (fTin = fTin) AND ((fTin - fTin) = (fTin - fTin))              (* 室内温 NaN 自反 + Inf 差判闸（边界④） / Indoor NaN and Inf gate *)
         AND (fTout = fTout) AND ((fTout - fTout) = (fTout - fTout));   (* 室外温 NaN 自反 + Inf 差判闸 / Outdoor NaN and Inf gate *)
tonPurge(IN := (_eState = E_DL_NfpState.ePurge), PT := tPurgeMax);      (* 吹扫超时：相位闸 + 无条件调用（边界②） / Purge timeout *)
tonCool(IN := (_eState = E_DL_NfpState.eHoldout), PT := tCooldown);     (* 冷却驻留：相位闸 + 无条件调用（边界②） / Cooldown timer *)

(* —— 段 1：单拍量预清零（R107） —— *)
bPurgeCmd := FALSE;                                      (* 吹扫命令出口预清（派生拍覆盖） / Purge command preset *)
bHoldout := FALSE;                                       (* 冷却指示出口预清 / Cooldown preset *)

(* —— 段 2：复位沿处理（作用域：清故障 + 清传感器锁存 + 迁 eIdle，R283 逐项声明） —— *)
IF rtReset.Q THEN
    _bFault := FALSE;                                    (* 清故障锁存 / Clear fault *)
    _eCause := E_DL_NfpCause.eNone;                      (* 清成因 / Clear cause *)
    bSensorBad := FALSE;                                 (* 清传感器失效锁存 / Clear sensor latch *)
    _bCoolDone := TRUE;                                  (* 冷却完成回 TRUE（复位即放行首轮） / Cooldown done reset *)
    _bDropOk := FALSE;                                   (* 清达标锁存 / Clear drop latch *)
    _eState := E_DL_NfpState.eIdle;                      (* 迁未吹扫相 / Back to idle *)
END_IF

(* —— 段 3：组态故障锁存（锁存至复位沿，R189） —— *)
IF _bCfgBad AND NOT _bFault THEN
    _bFault := TRUE;                                     (* 锁存故障位 / Latch fault *)
    _eCause := E_DL_NfpCause.eCfgIllegal;                (* 成因：组态非法 / Cause illegal config *)
    _eState := E_DL_NfpState.eFault;                     (* 同步迁故障相 / Migrate to fault *)
END_IF

(* —— 段 4：CASE 主状态机（ELSE 兜底迁 eFault，红线 6） —— *)
CASE _eState OF
    E_DL_NfpState.eIdle:                                 (* 未吹扫：出口确定值 / Idle *)
        bPurgeCmd := FALSE;                              (* 失能吹扫命令确定 FALSE / Disabled command false *)
        bHoldout := FALSE;                               (* 失能冷却指示 FALSE / Disabled holdout false *)
        IF bEnable AND NOT _bFault AND _bCoolDone AND _bFin              (* 使能 + 冷却窗满（边界⑤）+ 温度有限 / Entry preconditions *)
           AND bWindow AND bFanAllow                                     (* 日历窗 + 风机允许（边界①） / Window and fan permit *)
           AND (fTout < fTin - fDelta) THEN                              (* 室外低温差闸（边界①） / Outdoor cool delta *)
            _fTinStart := fTin;                          (* 迁入拍室内温快照（温降基准） / Indoor snapshot *)
            _bDropOk := FALSE;                           (* 清达标锁存（新一轮） / Clear drop latch *)
            _bCoolDone := FALSE;                         (* 冷却窗未满（退出后重计） / Cooldown not done *)
            _eState := E_DL_NfpState.ePurge;             (* 进入吹扫相 / Enter purging *)
        END_IF
    E_DL_NfpState.ePurge:                                 (* 吹扫相：达标/超时/降级三出口 / Purging *)
        bPurgeCmd := TRUE;                                (* 吹扫命令出口 / Purge command *)
        IF NOT bEnable OR NOT bWindow OR NOT bFanAllow OR NOT _bFin THEN   (* 前置消失或传感器失效（安全侧降级，边界④） / Preconditions lost *)
            IF NOT _bFin THEN
                bSensorBad := TRUE;                      (* 传感器失效锁存（复位沿清，边界④） / Sensor bad latch *)
                _eCause := E_DL_NfpCause.eSensorBad;     (* 成因：传感器失效 / Cause sensor bad *)
            END_IF
            _eState := E_DL_NfpState.eHoldout;           (* 降级入冷却驻留（安全侧不维持） / To cooldown *)
            _bDropOk := FALSE;                           (* 清达标锁存 / Clear drop latch *)
        ELSE
            IF (_fTinStart - fTin) >= fDropTgt THEN      (* 温降达标上阈（差值直比，边界③） / Drop reached upper *)
                _bDropOk := TRUE;                        (* 达标锁存 / Drop latch *)
            END_IF
            IF _bDropOk AND ((_fTinStart - fTin) < (fDropTgt - fDropHys)) THEN   (* 跌破迟滞下带才解除达标（边界③） / Release below band *)
                _bDropOk := FALSE;                       (* 解除达标 / Drop release *)
            END_IF
            IF _bDropOk OR tonPurge.Q THEN               (* 达标或超时退出 / Drop or timeout exit *)
                _eState := E_DL_NfpState.eHoldout;       (* 入冷却驻留窗（边界⑤） / To cooldown *)
                _bDropOk := FALSE;                       (* 清达标锁存 / Clear drop latch *)
            END_IF
        END_IF
    E_DL_NfpState.eHoldout:                              (* 冷却驻留相：窗满回未吹扫 / Cooldown *)
        bHoldout := TRUE;                                (* 冷却指示出口 / Cooldown indicator *)
        bPurgeCmd := FALSE;                              (* 冷却相吹扫命令确定 FALSE / Purge command false *)
        IF tonCool.Q THEN
            _bCoolDone := TRUE;                          (* 冷却窗满放行（边界⑤） / Cooldown done *)
            _eState := E_DL_NfpState.eIdle;              (* 回未吹扫相 / Back to idle *)
        END_IF
    E_DL_NfpState.eFault:                                (* 故障相：冻结保持，仅复位沿出 / Fault *)
        ;                                                (* 锁存回放（R28） / Replay from latch *)
    ELSE                                                 (* 非法相位兜底迁安全态 / Illegal phase fallback *)
        _eState := E_DL_NfpState.eFault; _bFault := TRUE;    (* 迁故障相 + 同步锁存 / To fault and latch *)
        _eCause := E_DL_NfpCause.ePhaseBad;              (* 成因：非法相位 / Cause illegal phase *)
END_CASE

(* —— 段 5：出口映射（bError/eState 同源，R191） —— *)
bError := _bFault;                                       (* 故障标志镜像 / Fault flag mirror *)
eState := _eState;                                       (* 状态出口 / State outlet *)
eCause := _eCause;                                       (* 成因出口 / Cause outlet *)
END_FUNCTION_BLOCK

(* ---- FB_DL_NightPurgeCtrl.st ---- *)
(*==============================================================================
 * 组件名称 (Component)  : FB_DL_NightPurgeCtrl
 * 所属子库 (Sublibrary) : DL_Process
 * 前缀     (Prefix)     : FB_DL_
 * 当前版本 (Version)    : 1.0.1
 * 兼容性   (Platform)   : CODESYS 3.5 / TwinCAT 3 / 汇川 InoProShop / Schneider
 *                         Machine Expert；纯 IEC 61131-3（第 3 版），
 *                         仅依赖标准库 TON 与库内 FC_DL_VaporPressureSat，
 *                         零厂商方言
 * 作者     (Author)     : 道莅代码库 · PLC编程专家（R31）
 * 开源溯源 (Origin)     : 夜间通风/免费冷却公开控制语义（T1-2 ROOM_CONTROL
 *                         族待挖子项），道莅 clean-room 防御性实现，
 *                         未复制任何外部源码行
 * 功能描述 (Function)   : 夜间吹扫顺控件（降温除湿侧方向写死，不出加热吹扫
 *                         变体）。三判据同时成立进入：无人员占用 + 室外比
 *                         室内凉（带死区）+ 室外绝对湿度不高于室内。窗时到
 *                         或判据失效退出；退出后经冷却时长抑制防频启。
 *                         Magnus-Tetens 饱和压常数唯一属主为库内
 *                         FC_DL_VaporPressureSat，本件只调用不内联公式。
 * 码位     (Codes)      : 16#0005_0094 信息级：温湿度非有限保持现状、
 *                         冷却期吹扫请求被拒、相对湿度越域已钳位（不置 bError）
 *                         16#0005_0095~0098 故障级保留未启用（本轮无故障级条件，
 *                         码表与实现对齐，不虚声明）
 * 边界防错 (Boundary)   : 1 温湿度非有限（x<>x 自反判加幅值界）保持现状+信息码；
 *                         2 相对湿度先钳 0..100 再参与换算；
 *                         3 TON 每拍无条件刷新，条件经入参传递；
 *                         4 CASE 带 ELSE 锁安全侧（不吹扫）；
 *                         5 饱和压调用失败按数据无效保持现状。
 * 规格偏离 (Deviation)   : 1 规格时戳类型 DTL 为平台扩展，改用 IEC 标准
 *                         DATE_AND_TIME（跨平台红线裁定），本轮判据不消费该
 *                         引脚，仅作观测时戳保留契约；
 *                         2 规格枚举名 E_DL_PurgeState 属主为库内
 *                         FB_DL_InertPurgeSeq（氮气置换语义），跨域语义不
 *                         复用，改立本文件私有枚举 E_DL_NightPurgeState。
 * 修订历史 (Revision)   : 2026-11-18 v1.0.0 首版入库（R31 · 阶段三 · 序 4）
 *                         2026-11-23 v1.0.1 R73 补 bValid 回执：段 3 两处饱和压
 *                         调用补收 bValid 局部回执，回执无效并入既有 bSat*Ok
 *                         拒绝语义（数据无效合取路径），契约不变
 *==============================================================================*)

(*------------------------------------------------------------------------------
 * 枚举: E_DL_NightPurgeState（归属本功能块，同文件发布，全库唯一属主）
 * 含义: 夜间吹扫（降温除湿侧）顺控状态，成员与 CASE 标签双向完备。
 *----------------------------------------------------------------------------*)
TYPE E_DL_NightPurgeState :
(
    eIdle     := 0,    // 待机：判据未齐或未使能 / Idle, criteria not met or disabled
    ePurging  := 10,   // 吹扫中：请求输出置位 / Purging, request output active
    eCooldown := 20,   // 冷却抑制：退出后重启抑制 / Cooldown, restart suppression after exit
    eFault    := 99    // 故障兜底：非法状态拦截 / Fault fallback, illegal state catch
);
END_TYPE

(*==============================================================================
 * 功能块: FB_DL_NightPurgeCtrl
 * 调用约定: 每个扫描周期无条件调用一次；实例状态全部驻留于私有变量。
 *==============================================================================*)
FUNCTION_BLOCK FB_DL_NightPurgeCtrl
VAR_INPUT
    bEn       : BOOL := FALSE;        // 使能 / Enable flag
    dtNow     : DT   := DT#1970-01-01-00:00:00; // 观测时戳（保留契约，本轮不消费）/ Observation timestamp, reserved
    fTOut     : REAL := 25.0;         // 室外温度 [摄氏度] / Outdoor temperature [degC]
    fTIn      : REAL := 25.0;         // 室内温度 [摄氏度] / Indoor temperature [degC]
    fRhOut    : REAL := 50.0;         // 室外相对湿度 [百分数] / Outdoor relative humidity [%]
    fRhIn     : REAL := 50.0;         // 室内相对湿度 [百分数] / Indoor relative humidity [%]
    fTDead    : REAL := 1.0;          // 温差判据死区 [摄氏度] / Temperature deadband [degC]
    tPurgeWin : TIME := T#60M;        // 吹扫窗口时长 [ms] / Purge window duration [ms]
    tCooldown : TIME := T#30M;        // 冷却抑制时长 [ms] / Cooldown suppression duration [ms]
    bOcc      : BOOL := FALSE;        // 人员占用信号 / Occupancy signal
END_VAR
VAR_OUTPUT
    bPurgeReq : BOOL;                 // 吹扫请求输出 / Purge request output
    eState    : E_DL_NightPurgeState; // 顺控当前状态 / Current sequence state
    uErrorId  : UDINT;                // 信息级码，0 = 无信息 / Info code, 0 = none
END_VAR
VAR
    tonWin    : TON;                  // 吹扫窗定时器，每拍无条件刷新 / Purge window timer, refreshed every scan
    tonCool   : TON;                  // 冷却抑制定时器，每拍无条件刷新 / Cooldown timer, refreshed every scan
    bCritOcc  : BOOL;                 // 判据一：无占用 / Criterion one: unoccupied
    bCritTemp : BOOL;                 // 判据二：室外比室内凉 / Criterion two: outdoor cooler
    bCritHum  : BOOL;                 // 判据三：室外绝对湿度不高于室内 / Criterion three: outdoor humidity not higher
    bCritOk   : BOOL;                 // 三判据合取 / All three criteria AND
    bDataOk   : BOOL;                 // 温湿度输入有效性 / Input data validity
    fRhOutC   : REAL;                 // 钳位后室外湿度 [百分数] / Clamped outdoor humidity [%]
    fRhInC    : REAL;                 // 钳位后室内湿度 [百分数] / Clamped indoor humidity [%]
    fPwsOut   : LREAL;                // 室外饱和水汽压 [帕] / Outdoor saturation vapour pressure [Pa]
    fPwsIn    : LREAL;                // 室内饱和水汽压 [帕] / Indoor saturation vapour pressure [Pa]
    fAhOut    : REAL;                 // 室外绝对湿度 [克每立方米] / Outdoor absolute humidity [g per m3]
    fAhIn     : REAL;                 // 室内绝对湿度 [克每立方米] / Indoor absolute humidity [g per m3]
    bSatOutOk : BOOL;                 // 室外饱和压调用有效 / Outdoor saturation call valid
    bSatInOk  : BOOL;                 // 室内饱和压调用有效 / Indoor saturation call valid
    bRhClamp  : BOOL;                 // 湿度越域钳位标志 / Humidity clamp flag
    _bPwsValid: BOOL;                 // 饱和压属主件输出可用回执 / Saturation owner FC outputs-usable receipt
    _bPwsClamped : BOOL;    // 属主件钳位回执（本件不消费，仅契约全回执） / Owner clamp receipt (unused, full-receipt contract)
    _nPwsErr     : UDINT;   // 属主件错误码回执 / Owner error-code receipt
    _bPwsError   : BOOL;    // 属主件故障级回执 / Owner fault-flag receipt
END_VAR
VAR CONSTANT
    DL_NPC_FIN   : REAL  := 1.0E30;   // REAL 有限幅值判界 / REAL finiteness magnitude bound
    DL_NPC_AH_K  : REAL  := 2.1674;   // 绝对湿度换算系数 [克·帕每开尔文每立方米] / Absolute humidity factor [g Pa per K per m3]
    DL_NPC_T0    : REAL  := 273.15;   // 绝对温标偏移 [开尔文] / Absolute temperature offset [K]
    DL_NPC_RHMAX : REAL  := 100.0;    // 相对湿度域上限 [百分数] / Relative humidity upper bound [%]
END_VAR

// ---- 段 1｜定时器无条件刷新（红线：禁入条件分支）------------------------------
tonWin(IN := (eState = ePurging), PT := tPurgeWin);   // 吹扫窗计时按态断输入 / Window timer input per state
tonCool(IN := (eState = eCooldown), PT := tCooldown); // 冷却计时按态断输入 / Cooldown timer input per state

// ---- 段 2｜输入有效性与湿度钳位 ------------------------------------------------
bDataOk := (fTOut = fTOut) AND (fTIn = fTIn)
       AND (ABS(fTOut) < DL_NPC_FIN) AND (ABS(fTIn) < DL_NPC_FIN)
       AND (fRhOut = fRhOut) AND (fRhIn = fRhIn)
       AND (ABS(fRhOut) < DL_NPC_FIN) AND (ABS(fRhIn) < DL_NPC_FIN); // 温湿度四点有限 / Four inputs finite
fRhOutC := MIN(MAX(fRhOut, 0.0), DL_NPC_RHMAX);       // 室外湿度钳 0..100 / Clamp outdoor humidity
fRhInC  := MIN(MAX(fRhIn, 0.0), DL_NPC_RHMAX);        // 室内湿度钳 0..100 / Clamp indoor humidity
bRhClamp := (fRhOut < 0.0) OR (fRhOut > DL_NPC_RHMAX)
         OR (fRhIn < 0.0) OR (fRhIn > DL_NPC_RHMAX);  // 越域判定 / Out-of-range detection

// ---- 段 3｜饱和压查询：常数唯一属主 FC_DL_VaporPressureSat，只调用不内联 --------
bSatOutOk := FC_DL_VaporPressureSat(fTempC := REAL_TO_LREAL(fTOut),
               fPvSat => fPwsOut, bValid => _bPwsValid, bClamped => _bPwsClamped, eErr => _nPwsErr, bError => _bPwsError); // 室外饱和压查询 / Query outdoor saturation pressure
bSatOutOk := bSatOutOk AND _bPwsValid;                 // 输出可用回执并入既有拒绝语义 / Merge outputs-usable receipt into existing reject semantics
bSatInOk := FC_DL_VaporPressureSat(fTempC := REAL_TO_LREAL(fTIn),
               fPvSat => fPwsIn, bValid => _bPwsValid, bClamped => _bPwsClamped, eErr => _nPwsErr, bError => _bPwsError); // 室内饱和压查询 / Query indoor saturation pressure
bSatInOk := bSatInOk AND _bPwsValid;                   // 输出可用回执并入既有拒绝语义 / Merge outputs-usable receipt into existing reject semantics

// ---- 段 4｜绝对湿度换算：AH = 2.1674·pv/(273.15+T) [克每立方米] -----------------
IF bDataOk AND bSatOutOk AND bSatInOk AND ((fTOut + DL_NPC_T0) > 0.0) AND ((fTIn + DL_NPC_T0) > 0.0) THEN
    fAhOut := DL_NPC_AH_K * REAL_TO_LREAL(fRhOutC) / 100.0 * fPwsOut
            / (REAL_TO_LREAL(fTOut) + DL_NPC_T0);      // 室外绝对湿度 / Outdoor absolute humidity
    fAhIn  := DL_NPC_AH_K * REAL_TO_LREAL(fRhInC) / 100.0 * fPwsIn
            / (REAL_TO_LREAL(fTIn) + DL_NPC_T0);       // 室内绝对湿度 / Indoor absolute humidity
    bCritHum := fAhOut <= fAhIn;                       // 判据三：室外不高（降温除湿侧）/ Outdoor not higher
ELSE
    fAhOut  := 0.0;                                    // 异常路径确定值 / Deterministic fallback value
    fAhIn   := 0.0;                                    // 异常路径确定值 / Deterministic fallback value
    bCritHum := FALSE;                                 // 数据无效判据不成立 / Invalid data fails criterion
END_IF

// ---- 段 5｜判据装配 ------------------------------------------------------------
bCritOcc  := NOT bOcc;                                // 判据一：无占用 / Unoccupied
bCritTemp := (fTOut + fTDead) < fTIn;                 // 判据二：室外加死区仍低于室内 / Outdoor plus deadband still cooler
bCritOk   := bCritOcc AND bCritTemp AND bCritHum AND bDataOk
          AND bSatOutOk AND bSatInOk;                 // 合取含数据有效性 / AND with data validity

// ---- 段 6｜状态机（CASE 带 ELSE 锁安全侧不吹扫）--------------------------------
CASE eState OF
    eIdle:
        bPurgeReq := FALSE;                            // 待机不吹扫 / No purge in idle
        IF bEn AND bCritOk THEN
            eState := ePurging;                        // 三判据齐进入吹扫 / Criteria met, start purge
        END_IF
    ePurging:
        bPurgeReq := bEn;                              // 吹扫请求随使能 / Purge follows enable
        IF (NOT bEn) OR (NOT bCritOk) OR tonWin.Q THEN
            eState := eCooldown;                       // 判据失效或窗时到退入冷却 / Exit to cooldown
        END_IF
    eCooldown:
        bPurgeReq := FALSE;                            // 冷却期不吹扫 / No purge in cooldown
        IF bCritOk THEN
            uErrorId := 16#0005_0094;                  // 信息级：冷却期请求被拒 / Info: request rejected in cooldown
        END_IF
        IF tonCool.Q THEN
            eState := eIdle;                           // 冷却满回待机 / Cooldown elapsed, back to idle
        END_IF
    eFault:
        bPurgeReq := FALSE;                            // 故障态安全侧不吹扫 / Fault keeps purge off
        IF NOT bEn THEN
            eState := eIdle;                           // 撤使能自愈回待机 / Self-heal on disable
        END_IF
    ELSE
        eState := eFault;                              // 非法状态兜底 / Illegal state fallback
END_CASE

// ---- 段 7｜信息码装配（数据无效/钳位/冷却期拒绝共用信息级槽）--------------------
IF (NOT bDataOk) OR (NOT bSatOutOk) OR (NOT bSatInOk) THEN
    uErrorId := 16#0005_0094;                          // 信息级：非有限或查询无效保持现状 / Info: non-finite or invalid call, hold
ELSIF bRhClamp THEN
    uErrorId := 16#0005_0094;                          // 信息级：湿度越域已钳位 / Info: humidity clamped
END_IF
END_FUNCTION_BLOCK

(* ---- FB_DL_NightPurgeSeq.st ---- *)
(*
  ==================================================================
  组件名 Component  : FB_DL_NightPurgeSeq
  分类   Category   : DL_Process
  复杂度 Complexity  : cx5
  版本   Version    : 1.0.1
  功能   Purpose    : 夜间免费制冷吹扫顺控。三重判据全满足才执行：夜间时段窗
                      （tNow 与窗起点终点比较；跨午夜用年内序数法判跨日，
                      全路径无 MOD）+ 室内外温差闸（带 0.5 K 回差）+ 开窗
                      许可。执行中许可失效即回驻留（不中断置故障）；最小
                      执行时长防反复启停。与防冻族分工为（利用冷量）。
  来源   Source     : t1-oscat-building（借鉴 OSCAT Building ROOM_CONTROL 夜间
                      通风待挖子项的域语义，clean-room 自研实现，未复制
                      OSCAT 任何源码行）
  溯源   Origin     : IEC 61131-3 标准语义的道莅防御性实现；夜间免费制冷为
                      公开暖通空调节能语义。
  平台   Platform   : 纯 IEC 61131-3（Standard.library: TON / R_TRIG，无私有库）
  分工声明 Split     : 与 DL_Process 存量防冻族（FrostProtectFreeze 等）分工
                      ——防冻件防低温损害，本件利用夜间冷量节能预冷，方向相反；
                      时段窗时刻由调用方（PRG 层时钟同步）经 tNow 引脚传入，
                      本件不读系统时钟。
  作者   Author     : 道莅代码库 · PLC 编程专家（R57）
  ------------------------------------------------------------------
  边界 Boundary     :
                      一 温差闸回差 0.5 K 常量：进入用全阈值，退出减回差；
                      二 开窗许可失效：执行中即回驻留相（R191 显式声明，
                         不中断置故障），窗口命令安全侧关闭；
                      三 跨午夜时段窗用年内序数法（起点日与次日 +1 判跨日），
                         全路径无 MOD；
                      四 最小执行时长 tMinRun 防反复启停（执行相退出门控）；
                      五 夜窗结束（_bNight 变假）执行相立即退出，不受 tMinRun
                         门控（v1.0.1 偏离段声明：外因一次性事件不会抖振，
                         防止温差持续满足时把热空气灌进建筑）；
                      六 锁存解除路径 = bReset 上升沿（唯一路径，R188）；
                      七 无全局变量、无外部变量声明、无物理地址寻址。
  修订记录 Revision  :
    2026-11-21  v1.0.0  R57 首版（批 4 · 序号 20）
    2026-11-21  v1.0.1  R58 返修：执行相原退出条件只有三条，温差始终满足时
                        吹扫会持续到日间（违背利用夜间冷量的存在理由），段 6
                        新增第四条退出「NOT _bNight 夜窗末退出」，不受 tMinRun
                        门控；边界四→五重排，功能描述同步。
  ==================================================================
*)

TYPE E_DL_NpsPhase :
(
    eDwell := 0,  // 驻留：三判据评估 / dwelling, the triple criteria evaluated
    ePurge := 10, // 执行：开窗吹扫 / purging, the windows commanded
    eFault := 90  // 故障：成因锁存 / fault, the cause latched
);
END_TYPE

TYPE E_DL_NpsFault :
(
    eNone      := 0, // 无成因 / no cause
    eCfgBad    := 1, // 组态非法：温差阈值或序数越域（故障级，与 bError 配对）/ an illegal config
    eSensorBad := 2, // 温度非有限（故障级，与 bError 配对）/ a non finite temperature
    ePhaseBad  := 3  // 非法相位兜底（故障级，与 bError 配对）/ an illegal phase fallback
);
END_TYPE

FUNCTION_BLOCK FB_DL_NightPurgeSeq
VAR_INPUT
    bEnable     : BOOL := TRUE;      // 使能，失能即回驻留关窗 [-] / enable, disabling dwells and closes
    bReset      : BOOL := FALSE;     // 复位上升沿清锁存 [-] / reset rising edge clears the latch
    tNow        : TOD := T#00:00:00; // 当前时刻 [时刻]，由调用方时钟源传入 / the current time, fed by the caller clock source
    fToutC      : LREAL := 15.0;     // 室外温度实测 [摄氏度] / the outdoor temperature [degree celsius]
    fTinC       : LREAL := 26.0;     // 室内温度实测 [摄氏度] / the indoor temperature [degree celsius]
    fDiffOnK    : LREAL := 3.0;      // 温差闸进入阈值 [开尔文]，域 大于回差 / the diff entry threshold [kelvin], above the hysteresis
    bWinPermit  : BOOL := FALSE;     // 开窗许可（风雨 / 消防联锁给出）[-] / the window permit from the rain and fire interlocks
    tNightStart : TOD := T#22:00:00; // 夜间窗起点 [时刻] / the night window start [time of day]
    tNightEnd   : TOD := T#06:00:00; // 夜间窗终点 [时刻]，早于起点表跨午夜 / the night window end, earlier than the start means overnight
    nDayOfYear  : INT := 200;        // 年内序数日 [日]，域 1..366 / the day of year ordinal [day], one through three hundred sixty six
    tMinRun     : TIME := T#300S;    // 最小执行时长 [毫秒]，防反复启停 / the minimum run duration against hunting
END_VAR
VAR_OUTPUT
    bPurgeRun  : BOOL := FALSE; // 吹扫执行电平 [-] / the purge run level
    bWinCmd    : BOOL := FALSE; // 开窗命令输出（安全侧常闭）[-] / the window command outlet, normally closed
    bCondOk    : BOOL := FALSE; // 三判据满足预备指示 [-] / the criteria ready indicator
    ePhase     : E_DL_NpsPhase := E_DL_NpsPhase.eDwell; // 相位出口 [枚举] / the phase outlet
    eFault     : E_DL_NpsFault := E_DL_NpsFault.eNone; // 成因出口，锁存回放 [枚举] / the cause outlet replayed
    bError     : BOOL := FALSE; // 故障锁存标志 [-] / the fault latch flag
END_VAR
VAR
    rtReset  : R_TRIG; // 复位沿检测，段 0 无条件刷新 / the reset edge
    tonMinRun: TON;    // 最小执行窗，段 0 无条件刷新 / the minimum run window
    _ePhase  : E_DL_NpsPhase := E_DL_NpsPhase.eDwell; // 内部相位，CASE 唯一写入目标 / the internal phase
    _eFaulC  : E_DL_NpsFault := E_DL_NpsFault.eNone; // 故障级成因，锁存至复位沿 / the fault cause, latched
    _bFault  : BOOL := FALSE; // 故障锁存位 [-] / the fault latch bit
    _bInit   : BOOL := FALSE; // 首扫初始化完成标志（R310）/ the first scan flag
    _bInOk   : BOOL := FALSE; // 双温度有限 [-] / both temperatures finite
    _bCfgOk  : BOOL := FALSE; // 组态域内 [-] / the config inside the domain
    _bNight  : BOOL := FALSE; // 当拍处于夜间窗 [-] / inside the night window this scan
    _bArmed  : BOOL := FALSE; // 跨午夜窗 armed 标记（起点日晚段已过）[-] / the overnight armed flag
    _nWinDay : INT := 0;      // 夜间窗起点日序数 [日] / the ordinal day the window opened
    _bDiffOk : BOOL := FALSE; // 温差闸回差锁存 [-] / the diff hysteresis latch
END_VAR
VAR CONSTANT
    DL_NP_DIFF_HYST : LREAL := 0.5; // 温差闸回差 [开尔文]（边界一）/ the diff hysteresis [kelvin]
    DL_NP_DOY_MAX   : INT := 366;   // 年内序数上界 [日] / the ordinal upper bound [day]
END_VAR

// 段 0｜定时器与沿检测无条件周期刷新（禁入分支）/ segment 0, the unconditional refresh
rtReset(CLK := bReset); // 复位沿 / the reset edge
tonMinRun(IN := (_ePhase = E_DL_NpsPhase.ePurge) AND (NOT _bFault), PT := tMinRun); // 最小执行窗，IN 串执行相闸 / the minimum run gated by the purge phase

// 段 1｜首扫初始化（R310）/ segment 1, the first scan
IF NOT _bInit THEN // 首扫一拍 / the first scan
    _bInit := TRUE; // 置首扫标志 / raise the flag
END_IF

// 段 2｜复位沿作用域：清锁存 / 清跨日标记 / 迁驻留（三项逐项声明）/ segment 2, the reset edge scope
IF rtReset.Q THEN // 复位沿 / the reset edge
    _bFault := FALSE; // 作用域一：清故障锁存 / scope one, clear the fault latch
    _eFaulC := E_DL_NpsFault.eNone; // 作用域一：清成因 / scope one, clear the cause
    _bArmed := FALSE; // 作用域二：清跨日 armed 标记 / scope two, clear the armed flag
    _nWinDay := 0; // 作用域二：清起点日序数 / scope two, clear the opening ordinal
    _ePhase := E_DL_NpsPhase.eDwell; // 作用域三：迁驻留相 / scope three, back to dwell
END_IF

// 段 3｜组态与输入域闸（R151 全覆盖）/ segment 3, the configuration and input gates
_bInOk := (fToutC = fToutC) AND ((fToutC - fToutC) = (fToutC - fToutC)) AND (fTinC = fTinC) AND ((fTinC - fTinC) = (fTinC - fTinC)); // 双温度有限双判据 / the dual temperature finiteness
_bCfgOk := (fDiffOnK > DL_NP_DIFF_HYST) AND (fDiffOnK = fDiffOnK) AND (nDayOfYear >= 1) AND (nDayOfYear <= DL_NP_DOY_MAX) AND (tMinRun > T#0S) AND (tNightStart <> tNightEnd); // 温差阈值 / 序数 / 最小时长 / 零长窗域判定（起点=终点判零长窗非法，R253）/ the threshold, ordinal, duration and zero length window verdicts
IF (NOT _bInOk) OR (NOT _bCfgOk) THEN // 输入缺陷或组态非法 / a defect or an illegal config
    IF NOT _bFault THEN // 未锁存才迁移 / migrate only while unlatched
        _bFault := TRUE; // 置故障锁存 / raise the fault latch
        IF NOT _bInOk THEN // 传感失效优先归因（R190）/ the sensor failure first
            _eFaulC := E_DL_NpsFault.eSensorBad; // 传感成因 / the sensor cause
        ELSE // 组态非法 / the illegal config
            _eFaulC := E_DL_NpsFault.eCfgBad; // 组态成因 / the config cause
        END_IF
        _ePhase := E_DL_NpsPhase.eFault; // 迁故障相 / migrate to fault
    END_IF
END_IF

// 段 4｜夜间时段窗判定（序数法判跨日，无 MOD，边界三）/ segment 4, the night window by the ordinal method
IF tNightStart < tNightEnd THEN // 同日窗路径（相等已由段 3 组态闸判非法，R253）/ the same day window path, equality judged illegal by segment three
    _bNight := (tNow >= tNightStart) AND (tNow <= tNightEnd); // 起点终点夹逼 / the span containment
    _bArmed := FALSE; // 同日窗不涉跨日 / no overnight involved
ELSE // 跨午夜窗路径 / the overnight window path
    IF tNow >= tNightStart THEN // 晚段：窗开启并记录起点日序数 / the evening segment, the window opens
        _bNight := TRUE; // 窗内 / inside
        _bArmed := TRUE; // 置 armed / arm
        _nWinDay := nDayOfYear; // 记起点日序数 / record the opening ordinal
    ELSIF tNow <= tNightEnd THEN // 早段：仅起点日或次日有效（序数法判跨日）/ the morning segment, the opening day or the next day only
        _bNight := _bArmed AND ((nDayOfYear = _nWinDay) OR (nDayOfYear = _nWinDay + 1)); // 序数法判跨日 / the ordinal cross day verdict
    ELSE // 白天空窗段 / the daytime gap
        _bNight := FALSE; // 窗外 / outside
        _bArmed := FALSE; // 清 armed / disarm
    END_IF
END_IF

// 段 5｜温差闸回差锁存（边界一）/ segment 5, the diff hysteresis latch
IF (fTinC - fToutC) > fDiffOnK THEN // 进入判据（全阈值）/ the entry with the full threshold
    _bDiffOk := TRUE; // 置温差锁存 / raise the diff latch
ELSIF (fTinC - fToutC) < (fDiffOnK - DL_NP_DIFF_HYST) THEN // 退出判据（减回差）/ the exit minus the hysteresis
    _bDiffOk := FALSE; // 清温差锁存 / clear the diff latch
END_IF

// 段 6｜相位机：ENUM + CASE，含 ELSE 非法相位兜底（R128）/ segment 6, the phase machine
CASE _ePhase OF

E_DL_NpsPhase.eDwell: // 驻留相：三判据齐全才执行 / the dwell phase, all three criteria start the purge
    IF NOT bEnable THEN // 失能 / disabled
        _ePhase := E_DL_NpsPhase.eDwell; // 停摆驻留 / dwell
    ELSIF _bNight AND _bDiffOk AND bWinPermit AND (NOT _bFault) THEN // 三判据齐全（时段 + 温差 + 许可）/ the triple criteria met
        _ePhase := E_DL_NpsPhase.ePurge; // 迁执行相 / migrate to purge
    END_IF

E_DL_NpsPhase.ePurge: // 执行相：退出条件 ≥4（失能 / 许可失效 / 夜窗结束 / 温差退出且最小时长满足，边界二一四五）/ the purge phase, at least four exit conditions
    IF NOT bEnable THEN // 失能 / disabled
        _ePhase := E_DL_NpsPhase.eDwell; // 回驻留相 / back to dwell
    ELSIF NOT bWinPermit THEN // 许可失效即回驻留，不中断置故障（边界二）/ the permit lost returns to dwell
        _ePhase := E_DL_NpsPhase.eDwell; // 回驻留相 / back to dwell
    ELSIF NOT _bNight THEN // 夜窗结束退出：外因一次性事件，不受 tMinRun 门控（边界五，v1.0.1）/ the night window end exits without the minimum gate
        _ePhase := E_DL_NpsPhase.eDwell; // 回驻留相 / back to dwell
    ELSIF (NOT _bDiffOk) AND tonMinRun.Q THEN // 温差退出且最小时长已满足（边界一四）/ the diff exit with the minimum met
        _ePhase := E_DL_NpsPhase.eDwell; // 回驻留相 / back to dwell
    END_IF

E_DL_NpsPhase.eFault: // 故障相：成因锁存，等复位沿；窗口命令安全侧关闭 / the fault phase, the command closed on the safe side
ELSE // 非法相位兜底（R128）/ the illegal phase fallback
    _bFault := TRUE; // 置故障锁存 / raise the fault latch
    _eFaulC := E_DL_NpsFault.ePhaseBad; // 故障级成因（R45 配对 bError）/ the fault cause
    _ePhase := E_DL_NpsPhase.eFault; // 迁故障相 / migrate to fault
END_CASE

// 段 7｜统一出口 / segment 7, the unified outlet
bPurgeRun := (_ePhase = E_DL_NpsPhase.ePurge) AND (NOT _bFault); // 执行电平 / the run level
bWinCmd := bPurgeRun; // 开窗命令与执行同源（安全侧常闭）/ the command shares the run source
bCondOk := _bNight AND _bDiffOk AND bWinPermit AND bEnable AND (NOT _bFault); // 预备指示 / the ready indicator
ePhase := _ePhase; // 相位出口单点映射 / the phase outlet
IF _bFault THEN // 故障锁存优先 / the fault latch first
    eFault := _eFaulC; // 成因锁存回放（R152）/ the cause replayed
ELSE // 无锁存 / no latch
    eFault := E_DL_NpsFault.eNone; // 无成因 / no cause
END_IF
bError := _bFault; // 故障标志与锁存位同源 / the flag shares the latch
END_FUNCTION_BLOCK

(* ---- FB_DL_NitrideFurnaceAmmoniaPurge.st ---- *)
(*==============================================================================
 * 组件名称 (Component)  : FB_DL_NitrideFurnaceAmmoniaPurge
 * 所属子库 (Sublibrary) : DL_Process
 * 归属目录 (Directory)  : C:\Library\DL_Process
 * 当前版本 (Version)    : 1.0.0
 * 分类/来源标签         : 功能块（FUNCTION_BLOCK）· 热处理工艺 · 氮化炉氨吹扫顺控
 *                         industry-pool / heat-treatment / nitriding / purge-seq
 * 兼容性   (Platform)   : CODESYS 3.5 / TwinCAT 3 / 汇川 InoProShop / 施耐德
 *                         Machine Expert；仅用 Standard.library 的 TON / ABS
 * 溯源声明 (Provenance) : 道莅自研 clean-room——只借公开规范条款与工程惯例，零代码行复制。
 * 功能一句话 (Summary)  : 氮化炉氨吹扫两段顺控：大流量吹扫 + 小流量置换，
 *                         氨分解率与残氨双判据，残氨排放联锁超限即中止。
 *
 * 功能描述 (Function)   : 六相状态机：待机/预检/一段吹扫/二段置换/合格判定/
 *                         中止保持。预检校验分解率与残氨数据有效；一段按
 *                         时限大流量吹扫，二段按时限小流量置换；任一相残氨
 *                         超联锁阈立即转中止保持（保守方向：氨阀关、氮阀
 *                         关、排放风机停），分解率域外或非有限同样中止；
 *                         两段时限全部走完且残氨合格转合格判定（信息级）。
 *                         中止保持仅撤使能或重新起动指令可解除。
 * 与既有件边界 (Boundary): 本件只编排吹扫阀组与排放风机，不控炉温；
 *                         氨分解率分析仪信号由引脚注入。
 * 码位说明 (Codes)      : 信息 16#0006_302D 吹扫合格完成
 *                         故障 16#0006_302E 输入非有限，保守中止
 *                         故障 16#0006_302F 残氨超排放联锁阈，中止保持
 *                         故障 16#0006_3030 分解率域外（小于 0 或大于 100）
 *                         段 16#06_0_2D~31 首槽信息级、次槽起故障级。
 * 依赖说明 (Depends)    : 无 DL_ 内部依赖；仅 Standard.library 的 TON / ABS。
 * 红线自检 (Redline)    : 零全局依赖 ｜ 零 VAR_EXTERNAL ｜ 零 %I/%Q（阀组引脚）
 *                         NaN/Inf 精确判据拦截 ｜ 浮点比较带 fEps 容差
 *                         ENUM 配 CASE 且 ELSE 兜底 ｜ TON 每周期无条件刷新
 *                         全变量双语同行注释 ｜ 安全联锁最高优先、保守失败方向
 * 修订历史 (Revision)   : 2026-11-18  v1.0.0  首版入库（R32 · 批 4）
 *============================================================================*)

FUNCTION_BLOCK FB_DL_NitrideFurnaceAmmoniaPurge
VAR_INPUT
    bRun       : BOOL;                    // 顺控使能，假则中止保持清故障 / Enable, FALSE aborts and clears
    bStart     : BOOL;                    // 起动指令 [事件]，待机相起动 / Start command
    fDissocPct : LREAL;                   // 氨分解率 [％]，域 0 到 100 / Ammonia dissociation percent
    fNh3Ppm    : LREAL;                   // 残氨浓度 [ppm] / Residual ammonia ppm
    fNh3IlkPpm : LREAL := 1000.0;         // 残氨排放联锁阈 [ppm] / Emission interlock threshold
    fNh3OkPpm  : LREAL := 200.0;         // 吹扫合格残氨阈 [ppm] / Purge pass threshold
    tStage1S   : TIME  := T#20M;          // 一段大流量吹扫时限 [s] / Stage 1 duration
    tStage2S   : TIME  := T#10M;          // 二段小流量置换时限 [s] / Stage 2 duration
    fEps       : LREAL := 1.0E-6;         // 浮点判零容差 [实数域] / Floating zero tolerance
END_VAR
VAR_OUTPUT
    oNh3Valve  : BOOL;                  // 氨阀输出 [引脚] / Ammonia valve output
    oN2Valve   : BOOL;                  // 氮阀输出 [引脚] / Nitrogen valve output
    oExhFan    : BOOL;                  // 排放风机输出 [引脚] / Exhaust fan output
    ePhase     : (ePhStandby := 0, ePhPrecheck := 1, ePhStage1 := 2, ePhStage2 := 3, ePhVerify := 4, ePhAbort := 5);  // 相枚举输出 / Phase output
    bDone      : BOOL;                  // 吹扫完成脉冲 [事件] / One-shot done pulse
    bError     : BOOL;                  // 故障标志，与故障码配对 / Fault flag paired with codes
    uErrorId   : UDINT;                 // 事件码，0 表示无事件 / Event code, zero means none
END_VAR
VAR
    _ePhase   : (ePhStandby := 0, ePhPrecheck := 1, ePhStage1 := 2, ePhStage2 := 3, ePhVerify := 4, ePhAbort := 5);   // 内部相 / Internal phase
    tonSt1    : TON;    // 一段时限定时器 [s]，每拍无条件刷新 / Stage 1 timer
    tonSt2    : TON;    // 二段时限定时器 [s]，每拍无条件刷新 / Stage 2 timer
    bSigOk    : BOOL;   // 分析数据有效标志 / Analyzer validity flag
    bStartEdge: BOOL;   // 起动沿暂存 / Start edge staging
    uCodeLatch: UDINT;  // 故障锁存码 [码] / Latched fault code
    uInfoCode : UDINT;  // 信息级单拍码 [码] / One-shot info code
    uPrevStart: BOOL;   // 上拍起动指令快照 [开关] / Previous start snapshot
END_VAR

(* 段 1｜定时器无条件刷新（红线 7）/ Timers refreshed unconditionally *)
tonSt1(IN := (_ePhase = ePhStage1) AND bRun, PT := tStage1S);    // 一段计时 / Stage 1 timing
tonSt2(IN := (_ePhase = ePhStage2) AND bRun, PT := tStage2S);    // 二段计时 / Stage 2 timing
bStartEdge := bStart AND (NOT uPrevStart);                       // 起动上升沿 / Start rising edge
uPrevStart := bStart;                                            // 快照更新 / Update the snapshot

(* 段 2｜分析数据有效性（每拍计算，判据门控挂状态量）/ Analyzer validity each scan *)
bSigOk := (fNh3Ppm = fNh3Ppm) AND (fDissocPct = fDissocPct)      // NaN 自反判据 / NaN reflexivity
          AND (ABS(fNh3Ppm) < 1.0E308) AND (ABS(fDissocPct) < 1.0E308)   // Inf 上限判据 / Inf limit
          AND (fDissocPct >= -fEps) AND (fDissocPct <= 100.0 + fEps);    // 分解率物理域 / Physical domain

(* 段 3｜最高优先级安全联锁（先于 CASE）：残氨超阈或数据无效即中止
 *      Highest-priority safety before the CASE: abort on interlock or bad data *)
IF (bRun AND bSigOk AND (fNh3Ppm > fNh3IlkPpm)) OR (bRun AND (NOT bSigOk) AND (_ePhase <> ePhStandby)) THEN
    _ePhase := ePhAbort;                // 拍 N 转中止保持 / To abort hold
    IF NOT bSigOk THEN
        uCodeLatch := 16#0006_302E;     // 故障级：数据非有限 / Fault: non-finite data
    ELSE
        uCodeLatch := 16#0006_302F;     // 故障级：残氨超联锁阈 / Fault: over interlock
    END_IF
END_IF
IF bRun AND bSigOk AND ((fDissocPct < -fEps) OR (fDissocPct > 100.0 + fEps)) THEN
    _ePhase := ePhAbort;                // 分解率域外中止 / Abort on out-of-domain dissociation
    uCodeLatch := 16#0006_3030;         // 故障级：分解率域外 / Fault: dissociation out of domain
END_IF

(* 段 4｜相状态机主分派（ENUM 配 CASE，ELSE 兜底）/ Phase dispatch with ELSE interception *)
CASE _ePhase OF

    ePhStandby:
        (* 本拍行为：阀组全关保守待机；使能与起动沿俱备拍 N+1 进预检 / Valves closed; arm on start edge *)
        oNh3Valve := FALSE;             // 关氨阀 / Close the ammonia valve
        oN2Valve := FALSE;              // 关氮阀 / Close the nitrogen valve
        oExhFan := FALSE;               // 停排放风机 / Stop the fan
        bDone := FALSE;                 // 完成脉冲清 / Clear the done pulse
        IF bRun AND bStartEdge THEN
            _ePhase := ePhPrecheck;     // 拍 N+1 进预检 / To precheck next scan
        END_IF

    ePhPrecheck:
        (* 本拍行为：数据有效即开阀起步；无效保守回待机 / Arm the valves when data valid *)
        IF NOT bSigOk THEN
            _ePhase := ePhAbort;        // 拍 N+1 中止 / To abort next scan
            uCodeLatch := 16#0006_302E; // 故障级：数据无效 / Fault: bad data
        ELSE
            oN2Valve := TRUE;           // 氮阀常开吹扫 / Nitrogen valve open
            oExhFan := TRUE;            // 排放风机开 / Fan on
            _ePhase := ePhStage1;       // 拍 N+1 进一段 / To stage 1 next scan
        END_IF

    ePhStage1:
        (* 本拍行为：氨阀开大流量吹扫，时限满转二段 / Big flow purge, transfer on time *)
        oNh3Valve := TRUE;              // 氨阀开 / Ammonia valve open
        oN2Valve := TRUE;               // 氮阀开 / Nitrogen valve open
        oExhFan := TRUE;                // 风机开 / Fan on
        IF NOT bRun THEN
            _ePhase := ePhAbort;        // 撤使能中止 / Disable aborts
        ELSIF tonSt1.Q THEN
            oNh3Valve := FALSE;         // 氨阀关进二段 / Close ammonia for stage 2
            _ePhase := ePhStage2;       // 拍 N+1 进二段 / To stage 2 next scan
        END_IF

    ePhStage2:
        (* 本拍行为：小流量氮置换，时限满转合格判定 / Small flow swap, transfer on time *)
        oNh3Valve := FALSE;             // 氨阀保持关 / Ammonia stays closed
        oN2Valve := TRUE;               // 氮阀开 / Nitrogen valve open
        oExhFan := TRUE;                // 风机开 / Fan on
        IF NOT bRun THEN
            _ePhase := ePhAbort;        // 撤使能中止 / Disable aborts
        ELSIF tonSt2.Q THEN
            _ePhase := ePhVerify;       // 拍 N+1 进合格判定 / To verify next scan
        END_IF

    ePhVerify:
        (* 本拍行为：残氨合格即完成（信息级），超合格阈但低于联锁阈转中止保守重来 / Verify *)
        oNh3Valve := FALSE;             // 阀组保持 / Valves held
        oN2Valve := TRUE;
        oExhFan := TRUE;
        IF fNh3Ppm <= fNh3OkPpm THEN
            oNh3Valve := FALSE;         // 全阀收 / Close all
            oN2Valve := FALSE;
            oExhFan := FALSE;
            bDone := TRUE;              // 完成脉冲（单拍）/ One-shot done
            uInfoCode := 16#0006_302D;  // 信息级：吹扫合格 / Info: purge passed
            _ePhase := ePhStandby;      // 拍 N+1 回待机 / To standby next scan
        ELSE
            _ePhase := ePhAbort;        // 拍 N+1 中止保守重来 / To abort, conservative retry
            uCodeLatch := 16#0006_302F; // 故障级：残氨未达合格阈 / Fault: residual over pass threshold
        END_IF

    ePhAbort:
        (* 本拍行为：保守中止三输出全关；撤使能或重新起动沿解除 / Conservative abort, all outputs closed *)
        oNh3Valve := FALSE;             // 全关保守方向 / All closed, conservative
        oN2Valve := FALSE;
        oExhFan := FALSE;               // 风机停防残氨扩散受控 / Fan off, controlled containment
        IF (NOT bRun) OR bStartEdge THEN
            uCodeLatch := 16#0000_0000; // 解除锁存（可达解除路径）/ Clear the latch, reachable reset
            _ePhase := ePhStandby;      // 拍 N+1 回待机 / To standby next scan
        END_IF

ELSE
    oNh3Valve := FALSE;                 // 非法相全关保守 / Illegal phase, all closed
    oN2Valve := FALSE;
    oExhFan := FALSE;
    _ePhase := ePhAbort;                // 拦截进中止 / Intercept to abort
    uCodeLatch := 16#0006_302E;         // 故障：相越界 / Fault: phase out of range
END_CASE

(* 段 5｜出口装配 / Exit assembly *)
ePhase := _ePhase;                      // 相枚举输出 / Phase output
bError := (uCodeLatch <> 16#0000_0000); // 故障锁存回放 / Latched fault replay
IF uCodeLatch <> 16#0000_0000 THEN
    uErrorId := uCodeLatch;             // 故障码优先 / Fault first
    uInfoCode := 16#0000_0000;
ELSE
    uErrorId := uInfoCode;              // 信息码单拍 / Info one shot
    uInfoCode := 16#0000_0000;
END_IF
END_FUNCTION_BLOCK

(* ---- FB_DL_OcvGradingBin.st ---- *)
(*
  FB_DL_OcvGradingBin  —  OCV 电压+内阻双判据分档与落料位决策 / OCV dual-criteria grading and bin decision
  分类 Category : DL_Process
  码位 Code     : 16#06_0_81
  版本 Version  : 1.0.0
  溯源 Source   : LGF Comparator 语义借鉴 · clean-room 实现，仅借分类/参数域/命名，未复制源码
  功能 Function : 1) 电压 + 内阻双判据同时落窗才分档，档位带由组态表给定；
                  2) 档位阈值单调递增校验，倒置即冻结并报码（不静默容错）；
                  3) 电压或内阻为 NaN 时判「不可分档」，绝不落入最低档；目标档满仓时走避让档，无可用料仓则停线。
  边界 Boundary : ① 档位阈值单调递增校验（倒置即冻结 + 报码）；
                  ② 电压/内阻任一 NaN 时判「不可分档」而非落最低档（x <> x 自反判据）；
                  ③ 满仓档位无可用料仓时停线（bLineStop），不静默落最低档；
                  ④ 电压/内阻先过物理域闸，域外按不可分档处理。
  依赖 Depends  : None

  码表 Error codes（本件子码步进 16#10，避让邻件码位）:
    16#0002_0681 故障级：档位阈值倒置或档数越界（组态闸锁存，需 bReset 清除）
    16#0002_0691 故障级：档位下标越界（枚举兜底路径）
    16#0002_06A1 信息级：满仓避让已生效 / 无可用料仓（不置 bError）
*)

TYPE E_DL_OcvGradePhase :
(
    eIdle       := 0,   // 空闲待料 / Idle awaiting cell
    eGrading    := 10,  // 双判据分档中 / Grading in progress
    eGraded     := 20,  // 已落档 / Graded
    eNoBin      := 30,  // 满仓避让失败 / Bin avoidance failed
    eUngradable := 40,  // 不可分档 / Ungradable cell
    eFault      := 90   // 组态故障锁定 / Configuration fault locked
);
END_TYPE

FUNCTION_BLOCK FB_DL_OcvGradingBin
VAR_INPUT
    bEnable    : BOOL;                            // 总使能，FALSE 回空闲 / Master enable
    bStart     : BOOL;                            // 分档触发，上升沿取一次测量 / Trigger, rising edge latches one measurement
    bReset     : BOOL;                            // 复位，上升沿清锁存故障 / Reset, clears the latched fault
    fVoltV     : REAL;                            // 电芯开路电压 [V]，域 0.5~5.0 / Cell open-circuit voltage [V]
    fIrMohm    : REAL;                            // 电芯内阻 [mOhm]，域 0.1~500.0 / Cell internal resistance [mOhm]
    nBinCount  : INT := 1;                        // 档位总数 [档]，域 1~8 / Bin count, 1..8
    afVoltLo   : ARRAY[1..8] OF REAL;             // 各档电压下限 [V] / Per-bin voltage lower limit [V]
    afVoltHi   : ARRAY[1..8] OF REAL;             // 各档电压上限 [V] / Per-bin voltage upper limit [V]
    afIrLo     : ARRAY[1..8] OF REAL;             // 各档内阻下限 [mOhm] / Per-bin resistance lower limit [mOhm]
    afIrHi     : ARRAY[1..8] OF REAL;             // 各档内阻上限 [mOhm] / Per-bin resistance upper limit [mOhm]
    abBinFull  : ARRAY[1..8] OF BOOL;             // 各档料仓满标志 [开关] / Per-bin full flag
    nFallbackBin : INT := 0;                      // 避让档号，0 = 无避让档 / Fallback bin, 0 = none
    fEps       : REAL := 1.0E-6;                  // 浮点判零容差 [1] / Floating zero tolerance
END_VAR
VAR_OUTPUT
    nBinOut    : INT;                             // 落料档号 1..8，0 = 不分档 / Target bin 1..8, 0 = none
    bGraded    : BOOL;                            // 本拍完成分档（单拍脉冲）/ Graded this scan, single pulse
    bUngradable: BOOL;                            // 不可分档标志（保持型）/ Ungradable flag, held
    bLineStop  : BOOL;                            // 停线请求（无可用料仓）/ Line stop request
    bConfigFault : BOOL;                          // 组态故障标志 / Configuration fault flag
    bError     : BOOL;                            // 故障标志，与故障级码配对 / Fault flag paired with fault codes
    uErrorId   : UDINT;                           // 事件码，0 = 无事件 / Event code, 0 = none
    eStateOut  : E_DL_OcvGradePhase;              // 状态机当前态，段尾单点映射 / Phase mapped at tail
END_VAR
VAR
    _eState    : E_DL_OcvGradePhase := E_DL_OcvGradePhase.eIdle;  // 内部状态 / Internal state
    rtrStart   : R_TRIG;                          // 分档触发沿 / Grading trigger edge
    rtrReset   : R_TRIG;                          // 复位沿 / Reset edge
    bCfgOk     : BOOL;                            // 组态合法标志 / Configuration valid flag
    bMonoOk    : BOOL;                            // 单调递增校验标志 / Monotonicity valid flag
    bFinite    : BOOL;                            // 输入有限性标志 / Input finiteness flag
    bDomainOk  : BOOL;                            // 输入物理域标志 / Input physical domain flag
    nN         : INT;                             // 生效档数（钳位后）/ Effective bin count after clamping
    nI         : INT;                             // 档位循环下标 / Bin loop index
    nHit       : INT;                             // 命中档号暂存，0 = 未命中 / Hit bin, 0 = none
    nUse       : INT;                             // 最终使用档号 / Finally used bin
    fVoltLat   : REAL;                            // 触发当拍锁存的电压 [V] / Latched voltage [V]
    fIrLat     : REAL;                            // 触发当拍锁存的内阻 [mOhm] / Latched resistance [mOhm]
    bLatValid  : BOOL;                            // 锁存有效（触发后保持）/ Latched sample valid
    uFault     : UDINT;                           // 锁存故障码 / Latched fault code
    uInfo      : UDINT;                           // 信息级码 / Information code
END_VAR
VAR CONSTANT
    DL_OCV_BINMAX  : INT := 8;                    // 档位数组上界 [档] / Bin array upper bound
    DL_OCV_VMIN    : REAL := 0.5;                 // 电压物理域下限 [V] / Voltage domain low [V]
    DL_OCV_VMAX    : REAL := 5.0;                 // 电压物理域上限 [V] / Voltage domain high [V]
    DL_OCV_IRMIN   : REAL := 0.1;                 // 内阻物理域下限 [mOhm] / Resistance domain low [mOhm]
    DL_OCV_IRMAX   : REAL := 500.0;               // 内阻物理域上限 [mOhm] / Resistance domain high [mOhm]
END_VAR

(* === 段 0 · 实例刷新（无条件周期调用）=== *)
rtrStart(CLK := bStart);                          // 每拍刷新分档触发沿
rtrReset(CLK := bReset);                          // 每拍刷新复位沿

(* === 段 1 · 组态闸：档数域 + 阈值单调递增（倒置即锁存报码）=== *)
nN := nBinCount;                                  // 档数取用前先钳位，防数组越界
IF nN < 1 THEN
    nN := 1;
END_IF
IF nN > DL_OCV_BINMAX THEN
    nN := DL_OCV_BINMAX;
END_IF
bCfgOk := (nBinCount >= 1) AND (nBinCount <= DL_OCV_BINMAX);   // 档数越界即组态非法
bMonoOk := TRUE;                                  // 单调性先置真，逐档否决
FOR nI := 1 TO DL_OCV_BINMAX DO
    IF nI <= nN THEN
        bMonoOk := bMonoOk AND (afVoltHi[nI] > afVoltLo[nI])       // 单档电压上下限配比
                   AND (afIrHi[nI] >= afIrLo[nI]);                 // 单档内阻上下限配比
        IF nI > 1 THEN
            bMonoOk := bMonoOk AND (afVoltHi[nI] > afVoltHi[nI - 1]);   // 电压上沿严格单调递增
        END_IF
    END_IF
END_FOR
IF (NOT bCfgOk) OR (NOT bMonoOk) THEN
    uFault := 16#0002_0681;                       // 故障级：阈值倒置或档数越界，组态闸锁存
END_IF
IF rtrReset.Q AND bCfgOk AND bMonoOk THEN
    uFault := 16#0000;                            // 组态修正后复位沿解锁（故障码复位路径可达）
END_IF

(* === 段 2 · 输入域闸：NaN 用自反判据，域外按不可分档处理 === *)
bFinite := (fVoltV = fVoltV) AND (fIrMohm = fIrMohm)               // x <> x 自反判 NaN
           AND (ABS(fVoltV) < 1.0E30) AND (ABS(fIrMohm) < 1.0E30);  // 上限兜底判 Inf
bDomainOk := (fVoltV >= DL_OCV_VMIN) AND (fVoltV <= DL_OCV_VMAX)
             AND (fIrMohm >= DL_OCV_IRMIN) AND (fIrMohm <= DL_OCV_IRMAX);
IF rtrStart.Q THEN
    fVoltLat := fVoltV;                           // 触发沿锁存本次测量，分档期间不被刷新
    fIrLat := fIrMohm;                            // 内阻同步锁存
    bLatValid := TRUE;                            // 锁存有效
END_IF

(* === 段 3 · 主状态机（ENUM + CASE，含 ELSE 兜底）=== *)
CASE _eState OF
E_DL_OcvGradePhase.eIdle :
    nBinOut := 0;                                 // 未分档，档号 0
    bGraded := FALSE;                             // 分档脉冲复位（非置位型标志）
    bUngradable := FALSE;                         // 不可分档标志复位
    bLineStop := FALSE;                           // 停线请求复位
    IF uFault <> 16#0000 THEN
        _eState := E_DL_OcvGradePhase.eFault;     // 组态故障优先
    ELSIF rtrStart.Q THEN
        _eState := E_DL_OcvGradePhase.eGrading;   // 本拍进入分档相
    END_IF

E_DL_OcvGradePhase.eGrading :
    IF (NOT bFinite) OR (NOT bDomainOk) THEN
        bUngradable := TRUE;                      // 本拍行为：不可分档，绝不落最低档
        nBinOut := 0;
        uInfo := 16#0002_06A1;                    // 信息级：不可分档（不置 bError）
        _eState := E_DL_OcvGradePhase.eUngradable;
    ELSE
        nHit := 0;                                // 命中档号先清零
        FOR nI := 1 TO nN DO
            IF (fVoltLat >= afVoltLo[nI]) AND (fVoltLat <= afVoltHi[nI])
               AND (fIrLat >= afIrLo[nI]) AND (fIrLat <= afIrHi[nI]) THEN
                nHit := nI;                       // 双判据同时落窗才命中
                EXIT;
            END_IF
        END_FOR
        IF nHit = 0 THEN
            bUngradable := TRUE;                  // 双判据无交集：不可分档
            nBinOut := 0;
            _eState := E_DL_OcvGradePhase.eUngradable;
        ELSE
            nUse := nHit;                         // 默认落命中档
            IF abBinFull[nHit] THEN
                IF (nFallbackBin >= 1) AND (nFallbackBin <= nN) AND (NOT abBinFull[nFallbackBin]) THEN
                    nUse := nFallbackBin;         // 满仓避让到可用料仓
                    uInfo := 16#0002_06A1;        // 信息级：满仓避让生效
                ELSE
                    nUse := 0;                    // 无可用料仓
                    bLineStop := TRUE;            // 停线，禁止静默落最低档
                    uInfo := 16#0002_06A1;        // 信息级：无可用料仓
                    _eState := E_DL_OcvGradePhase.eNoBin;
                END_IF
            END_IF
            IF nUse >= 1 THEN
                nBinOut := nUse;                  // 落料档号输出
                bGraded := TRUE;                  // 置位型：完成脉冲，段尾不清零
                _eState := E_DL_OcvGradePhase.eGraded;
            END_IF
        END_IF
    END_IF

E_DL_OcvGradePhase.eGraded :
    bLatValid := FALSE;                           // 本拍行为：测量已消费，锁存失效
    _eState := E_DL_OcvGradePhase.eIdle;          // 转出：下一拍回空闲待料

E_DL_OcvGradePhase.eNoBin :
    bLineStop := TRUE;                            // 停线请求保持，直到人工处理
    IF rtrReset.Q THEN
        bLineStop := FALSE;                       // 复位沿解除停线（可到达的解除路径）
        uInfo := 16#0000;                         // 信息码同步清除
        _eState := E_DL_OcvGradePhase.eIdle;
    END_IF

E_DL_OcvGradePhase.eUngradable :
    IF rtrStart.Q THEN
        _eState := E_DL_OcvGradePhase.eGrading;   // 新料触发重新分档
    ELSIF rtrReset.Q THEN
        bUngradable := FALSE;                     // 复位沿清不可分档标志
        _eState := E_DL_OcvGradePhase.eIdle;
    END_IF

E_DL_OcvGradePhase.eFault :
    nBinOut := 0;                                 // 故障态不分档（安全侧）
    IF uFault = 16#0000 THEN
        _eState := E_DL_OcvGradePhase.eIdle;      // 故障已解锁则回空闲
    END_IF

ELSE
    _eState := E_DL_OcvGradePhase.eFault;         // 非法状态拦截
    nBinOut := 0;                                 // 安全侧档号
    uFault := 16#0002_0691;                       // 故障级：档位下标越界（枚举兜底路径）
END_CASE
IF NOT bEnable THEN
    _eState := E_DL_OcvGradePhase.eIdle;          // 失能最高优先回空闲
    nBinOut := 0;                                 // 档号随之为 0
    bLineStop := FALSE;                           // 失能时不停线
END_IF

(* === 段 4 · 输出映射与故障码汇总 === *)
bConfigFault := (uFault <> 16#0000);              // 组态故障标志
bError := (uFault <> 16#0000);                    // 故障标志仅由故障级码置位（R45 配对）
IF bError THEN
    uErrorId := uFault;                           // 故障级优先上报
ELSE
    uErrorId := uInfo;                            // 否则上报信息级码
END_IF
eStateOut := _eState;                             // 输出枚举段尾单点映射（N2 规则）
END_FUNCTION_BLOCK
